(* IEC 61131-3 sources: PLC-IsaVODE/PLC-IsaVODE/samples/plc-programs (part 8) *)

(* ---- 638-IRTRANS_SERVER.ST ---- *)
TYPE

  oscat_NW_BUF_SHORT : ARRAY [0..1407] OF BYTE;
  oscat_NW_BUF_LONG  : ARRAY [0..4095] OF BYTE;

  oscat_NETWORK_BUFFER_SHORT :
  STRUCT
    SIZE   : UINT;
    BUFFER : oscat_NW_BUF_SHORT;
  END_STRUCT;

  oscat_NETWORK_BUFFER :
  STRUCT
    SIZE   : UINT;
    BUFFER : oscat_NW_BUF_LONG;
  END_STRUCT;

END_TYPE

TYPE
  oscat_IP_FIFO128_DATA  : ARRAY [1..128] OF BYTE;
  oscat_Mailbox  : ARRAY [1..16] OF BYTE;

  oscat_IP_FIFO_DATA :
  STRUCT
	X       : oscat_IP_FIFO128_DATA; (* IP_ID FIFO Speicher          *)
	Y       : oscat_IP_FIFO128_DATA; (* IP_ID Z�hler                 *)
	ID      : BYTE;                  (* h�chste vergabene id         *)
	MAX_ID  : BYTE;                  (* maximal Anmeldungen pro ID   *)
    INIT    : BOOL;                  (* Initialisierung durchgef�hrt *)
	EMPTY   : BOOL;                  (* FIFO leer                    *)
	FULL    : BOOL;                  (* FIFO voll                    *)
	TOP     : INT;                   (* maximale anzahl in FIFO      *)
	NW      : INT;                   (* Schreibzeiger                *)
	NR      : INT;                   (* Lesezeiger                   *)
  END_STRUCT;

  oscat_IP_C:
  STRUCT
  	C_MODE:			BYTE;          		(*W Mode: TCP/UCP AKTIV/PASSIV                               *)
	C_PORT:         WORD;          		(*W Portnummer                                               *)
	C_IP:           DWORD;         		(*W IP-Adresse gepackt wwxxyyzz = www.xxx.yyy.zzz            *)
    C_STATE:        BYTE;          		(*R Verbindungsstatus ON/OFF + Flanke ON/OFF                 *)
	C_ENABLE:       BOOL;          		(*W Freigabe f�r Connect                                     *)
    R_OBSERVE:      BOOL;          		(*W Empfang ueberwachen                                      *)
    TIME_RESET:     BOOL;          		(*W Alle Timer ruecksetzen                                   *)
	ERROR:          DWORD;         		(*R vvwwxxyy (vv = CON_ERROR, ww = SEN_ERROR, xx = REC_ERROR *)
    FIFO:           oscat_IP_FIFO_DATA; (*I IP FIFO Struktur                                         *)
	MAILBOX:		oscat_Mailbox;		(*I Mailbox: Datenbereich f�r Bausteindatenaustausch         *)
  END_STRUCT;
END_TYPE

FUNCTION_BLOCK IRTRANS_SERVER_Block

	VAR_INPUT
		UDP_TCP :	BOOL;
	END_VAR

	VAR_OUTPUT
		S_ENABLE :	BOOL;
		R_ENABLE :	BOOL;
		ERROR :	DWORD;
	END_VAR

	VAR_IN_OUT
		IP_C :	oscat_IP_C;
		S_BUF :	oscat_NETWORK_BUFFER;
		R_BUF :	oscat_NETWORK_BUFFER;
	END_VAR

	VAR
		t :	TON;
	END_VAR

	IF NOT IP_C.C_ENABLE THEN
		IP_C.C_PORT := WORD#0;
		IP_C.C_IP := DWORD#00;
		IP_C.C_MODE := SEL(UDP_TCP,BYTE#5,BYTE#4);
		IP_C.C_ENABLE := TRUE;
		IP_C.R_OBSERVE := FALSE;
		IP_C.TIME_RESET := TRUE;
		S_BUF.SIZE := UINT#0;
		R_BUF.SIZE := UINT#0;
	END_IF;

	R_ENABLE := IP_C.C_STATE > BYTE#127;
	S_ENABLE := R_ENABLE AND (IP_C.MAILBOX[1] > BYTE#0 OR IP_C.C_MODE <> BYTE#5);
	ERROR := IP_C.ERROR;

	t(IN:= IP_C.ERROR > DWORD#0, PT:=T#5s);
	IF t.Q THEN
		IP_C.TIME_RESET := TRUE;
	END_IF;

END_FUNCTION_BLOCK

PROGRAM program0
	VAR
		UDP_TCP :	BOOL;
		S_ENABLE :	BOOL;
		R_ENABLE :	BOOL;
		ERROR :	DWORD;
		IP_C :	oscat_IP_C;
		S_BUF :	oscat_NETWORK_BUFFER;
		R_BUF :	oscat_NETWORK_BUFFER;

		func_block : IRTRANS_SERVER_Block;
	END_VAR
	func_block.UDP_TCP := UDP_TCP;
	func_block.IP_C := IP_C;
	func_block.S_BUF := S_BUF;
	func_block.R_BUF := R_BUF;

	func_block();
	S_ENABLE  := func_block.S_ENABLE;
	R_ENABLE  := func_block.R_ENABLE;
	ERROR  := func_block.ERROR;
	IP_C  := func_block.IP_C;
	S_BUF  := func_block.S_BUF;
	R_BUF  := func_block.R_BUF;

END_PROGRAM

CONFIGURATION Config0

  	RESOURCE Res0 ON PLC
    	TASK task0(INTERVAL := T#20ms,PRIORITY := 0);
    	PROGRAM instance0 WITH task0 : program0;
  	END_RESOURCE

END_CONFIGURATION

(* ---- 639-FT_PDT1.ST ---- *)
FUNCTION _REAL_TO_UDINT:UDINT
  VAR_INPUT
    X :	REAL;
  END_VAR

  IF REAL_TO_UDINT(0.5) = UDINT#1 THEN
    _REAL_TO_UDINT := REAL_TO_UDINT(x);
  ELSIF X > 0.0 THEN
    _REAL_TO_UDINT := REAL_TO_UDINT(x+0.5);
  ELSIF X < 0.0 THEN
    _REAL_TO_UDINT := REAL_TO_UDINT(x-0.5);
  ELSE
    _REAL_TO_UDINT := UDINT#0;
  END_IF;
END_FUNCTION

FUNCTION REAL_TO_TIME2:TIME
	VAR_INPUT
		IN :	REAL;
	END_VAR

	REAL_TO_TIME2 := DINT_TO_TIME(UDINT_TO_DINT(_REAL_TO_UDINT(IN)));
END_FUNCTION

FUNCTION_BLOCK T_PLC_US_Block
	VAR_OUTPUT
		T_PLC_US :	UDINT;
	END_VAR

	VAR_EXTERNAL
		PLC_TICKS_PER_SEC :	INT;
		PLC_SYS_TICK_CNT :	DINT;
	END_VAR

	VAR
		debug :	BOOL;
		N :	INT;
		Offset :	UDINT;
		temp :	DWORD := DWORD#1;
		mode :	BOOL;
		faktor :	UDINT;
		init :	BOOL;
		v_plc_ticks_per_sec :	UDINT;
		base :	UDINT := UDINT#1000000;
	END_VAR

	IF init = FALSE THEN
		v_plc_ticks_per_sec := INT_TO_UDINT(PLC_TICKS_PER_SEC);
		IF v_plc_ticks_per_sec = UDINT#1024 THEN
			faktor := UDINT#1000;
			mode := FALSE;
		ELSIF v_plc_ticks_per_sec > UDINT#0 THEN
			IF v_plc_ticks_per_sec <= base THEN
				faktor := base / v_plc_ticks_per_sec;
				mode := FALSE;
			ELSE
				faktor := v_plc_ticks_per_sec / base;
				mode := TRUE;
			END_IF;
		ELSE
			faktor := UDINT#1;
		END_IF;
		init := TRUE;
	END_IF;

	IF mode THEN
		T_PLC_US := DINT_TO_UDINT(PLC_SYS_TICK_CNT) / faktor;
	ELSE
		T_PLC_US := DINT_TO_UDINT(PLC_SYS_TICK_CNT) * faktor;
	END_IF;

	IF debug THEN
		T_PLC_US := (DWORD_TO_UDINT(SHL(UDINT_TO_DWORD(T_PLC_US),N) OR SHL(temp,N)) - UDINT#1) + Offset;
	END_IF;
END_FUNCTION_BLOCK

FUNCTION_BLOCK FT_DERIV
	VAR_INPUT
		IN :	REAL;
		K :	REAL := 1.0;
		RUN :	BOOL := TRUE;
	END_VAR

	VAR_OUTPUT
		OUT :	REAL;
	END_VAR

	VAR
		old :	REAL;
		tx :	UDINT;
		last :	UDINT;
		init :	BOOL;
		tc :	REAL;
		T_PLC_US :	T_PLC_US_Block;
	END_VAR

	T_PLC_US();
	tx:= T_PLC_US.T_PLC_US;
	tc := UDINT_TO_REAL(tx - last);

	IF NOT init THEN
		init := TRUE;
		old := in;
	ELSIF run AND tc > 0.0 THEN
		out := (in - old) / tc * 1000000.0 * K;
		old := in;
	ELSE
		out := 0.0;
	END_IF;

	last := tx;

	T_PLC_US();
	tx:= T_PLC_US.T_PLC_US;

	IF NOT init THEN
		init := TRUE;
	ELSIF run AND tx - last > UDINT#0 THEN
		out := (in - old) / UDINT_TO_REAL(tx - last) * 1000000.0 * K;
	ELSE
		out := 0.0;
	END_IF;
	old := in;
	last := tx;
END_FUNCTION_BLOCK

FUNCTION_BLOCK FT_PT1

	VAR_INPUT
		IN :	REAL;
		T :	TIME;
		K :	REAL := 1.0;
	END_VAR

	VAR_OUTPUT
		OUT :	REAL;
	END_VAR

	VAR
		last :	UDINT;
		tx :	UDINT;
		init :	BOOL;
		T_PLC_US :	T_PLC_US_Block;
	END_VAR

	T_PLC_US();
	tx:= T_PLC_US.T_PLC_US;

	IF NOT init OR T = t#0s THEN
		init := TRUE;
		out := K * in;
	ELSE
		out := out + (in * K - out) * UDINT_TO_REAL(Tx - last) / TIME_TO_REAL(T) * 1.0E-3;
		IF ABS(out) < 1.0E-20 THEN out := 0.0; END_IF;
	END_IF;
	last := tx;
END_FUNCTION_BLOCK

FUNCTION_BLOCK FT_PDT1_Block

	VAR_INPUT
		IN :	REAL;
		KP :	REAL := 1.0;
		TV :	REAL := 1.0;
		T1 :	REAL := 1.0;
	END_VAR

	VAR_OUTPUT
		Y :	REAL;
	END_VAR

	VAR
		diff :	FT_DERIV;
		_TP :	FT_PT1;
	END_VAR

	diff(IN := IN, K := TV);

	_tp(in := diff.out, T := REAL_TO_TIME2(T1));

	Y := KP * (_tp.out + IN);

END_FUNCTION_BLOCK

PROGRAM program0
	VAR
		IN :	REAL;
		KP :	REAL := 1.0;
		TV :	REAL := 1.0;
		T1 :	REAL := 1.0;

		Y :	REAL;
		func_block : FT_PDT1_Block;
	END_VAR
	func_block.IN :=IN;
	func_block.KP :=KP;
	func_block.TV :=TV;
	func_block.T1 :=T1;
	func_block();
	Y := func_block.Y;
END_PROGRAM

CONFIGURATION Config0

	VAR_GLOBAL
		PLC_TICKS_PER_SEC :	INT;
		PLC_SYS_TICK_CNT :	DINT;
	END_VAR

	RESOURCE Res0 ON PLC
		TASK task0(INTERVAL := T#20ms,PRIORITY := 0);
		PROGRAM instance0 WITH task0 : program0;
	END_RESOURCE

END_CONFIGURATION

(* ---- 640-BOILER.ST ---- *)
FUNCTION_BLOCK BOILER_Block

	VAR_INPUT
		T_UPPER :	REAL;
		T_LOWER :	REAL;
		PRESSURE :	BOOL := TRUE;
		ENABLE :	BOOL := TRUE;
		REQ_1 :	BOOL;
		REQ_2 :	BOOL;
		BOOST :	BOOL;
		T_UPPER_MIN :	REAL := REAL#50.0;
		T_UPPER_MAX :	REAL := REAL#60.0;
		T_LOWER_ENABLE :	BOOL;
		T_LOWER_MAX :	REAL := REAL#60.0;
		T_REQUEST_1 :	REAL := REAL#70.0;
		T_REQUEST_2 :	REAL := REAL#50.0;
		T_REQUEST_HYS :	REAL := REAL#5.0;
		T_PROTECT_HIGH :	REAL := REAL#80.0;
		T_PROTECT_LOW :	REAL := REAL#10.0;
	END_VAR

	VAR_OUTPUT
		HEAT :	BOOL;
		ERROR :	BOOL;
		STATUS :	BYTE;
	END_VAR

	VAR
		edge :	BOOL;
		boost_mode :	BOOL;
		flag_0 :	BOOL;
		flag_1 :	BOOL;
		flag_2 :	BOOL;
	END_VAR

	IF t_upper > t_protect_high THEN
		status := BYTE#1;
		heat := FALSE;
		error := TRUE;
	ELSIF t_upper < t_protect_low THEN
		status := BYTE#2;
		heat := TRUE;
		error := TRUE;
	ELSIF t_lower > T_protect_high AND t_lower_enable THEN
		status := BYTE#3;
		heat := FALSE;
		error := TRUE;
	ELSIF t_lower < t_protect_low AND t_lower_enable THEN
		status := BYTE#4;
		heat := TRUE;
		error := TRUE;
	ELSIF NOT pressure THEN
		status := BYTE#5;
		heat := FALSE;
		error := TRUE;
	ELSIF req_1 OR req_2 OR enable OR boost THEN
		error := FALSE;

		IF boost AND NOT edge AND t_upper < t_upper_max THEN
			status := BYTE#101;
			heat := TRUE;
			boost_mode := TRUE;
		ELSIF enable AND t_upper < T_upper_min THEN
			status := BYTE#102;
			heat := TRUE;
		ELSIF req_1 AND t_upper < T_request_1 THEN
			status := BYTE#103;
			heat := TRUE;
		ELSIF req_2 AND t_upper < t_request_2 THEN
			status := BYTE#104;
			heat := TRUE;
		END_IF;

		IF heat THEN
			IF (enable OR boost_mode) THEN
				flag_0 := TRUE;
				IF T_lower_enable AND T_lower > T_lower_max THEN
					flag_0 := FALSE;
					boost_mode := FALSE;
				ELSIF NOT T_lower_enable AND T_upper > T_upper_max THEN
					flag_0 := FALSE;
					boost_mode := FALSE;
				END_IF;
			ELSE
				flag_0 := FALSE;
			END_IF;
			flag_1 := (req_1 AND T_upper > T_request_1 + T_request_hys) AND req_1;
			flag_2 := (req_2 AND T_upper > T_request_2 + T_request_hys) AND req_2;

			heat := flag_0 OR flag_1 OR flag_2;
			IF heat = FALSE THEN status := BYTE#100; END_IF;
		END_IF;
	ELSE
		status := BYTE#100;
		heat := FALSE;
		error := FALSE;
	END_IF;
	edge := boost;

END_FUNCTION_BLOCK

PROGRAM program0
	VAR
		T_UPPER :	REAL;
		T_LOWER :	REAL;
		PRESSURE :	BOOL := TRUE;
		ENABLE :	BOOL := TRUE;
		REQ_1 :	BOOL;
		REQ_2 :	BOOL;
		BOOST :	BOOL;
		T_UPPER_MIN :	REAL := REAL#50.0;
		T_UPPER_MAX :	REAL := REAL#60.0;
		T_LOWER_ENABLE :	BOOL;
		T_LOWER_MAX :	REAL := REAL#60.0;
		T_REQUEST_1 :	REAL := REAL#70.0;
		T_REQUEST_2 :	REAL := REAL#50.0;
		T_REQUEST_HYS :	REAL := REAL#5.0;
		T_PROTECT_HIGH :	REAL := REAL#80.0;
		T_PROTECT_LOW :	REAL := REAL#10.0;
		HEAT :	BOOL;
		ERROR :	BOOL;
		STATUS :	BYTE;

		func_block : BOILER_Block;
	END_VAR
	func_block.T_UPPER := T_UPPER;
	func_block.T_LOWER := T_LOWER;
	func_block.PRESSURE := PRESSURE ;
	func_block.ENABLE    := ENABLE    ;
	func_block.REQ_1 := REQ_1;
	func_block.REQ_2 := REQ_2;
	func_block.BOOST := BOOST ;
	func_block.T_UPPER_MIN := T_UPPER_MIN ;
	func_block.T_UPPER_MAX    := T_UPPER_MAX    ;
	func_block.T_LOWER_ENABLE := T_LOWER_ENABLE;
	func_block.T_LOWER_MAX := T_LOWER_MAX;
	func_block.T_REQUEST_1 := T_REQUEST_1 ;
	func_block.T_REQUEST_2 := T_REQUEST_2 ;
	func_block.T_REQUEST_HYS    := T_REQUEST_HYS    ;
	func_block.T_PROTECT_HIGH := T_PROTECT_HIGH;
	func_block.T_PROTECT_LOW := T_PROTECT_LOW;

	func_block();
	HEAT  := func_block.HEAT;
	ERROR  := func_block.ERROR;
	STATUS  := func_block.STATUS;
END_PROGRAM

CONFIGURATION Config0
	RESOURCE Res0 ON PLC
		TASK task0(INTERVAL := T#20ms,PRIORITY := 0);
		PROGRAM instance0 WITH task0 : program0;
	END_RESOURCE
END_CONFIGURATION

(* ---- 641-RMP_SOFT.ST ---- *)
FUNCTION TIME_TO_UDINT2:UDINT
	VAR_INPUT
		X :	TIME;
	END_VAR

	TIME_TO_UDINT2 := DINT_TO_UDINT(TIME_TO_DINT(X));
END_FUNCTION

FUNCTION_BLOCK T_PLC_MS_block
	VAR_OUTPUT
		T_PLC_MS :	UDINT;
	END_VAR

	VAR_EXTERNAL
		PLC_TICKS_PER_SEC :	INT;
		PLC_SYS_TICK_CNT :	DINT;
	END_VAR

	VAR
		debug :	BOOL;(*Debug-Mode ON / OFF*)
		N :	INT;(*Debug-Faktor*)
		Offset :	UDINT;(*Debug-Offset*)
		temp :	DWORD := DWORD#1;(*Debug-Offset*)
		mode :	BOOL;(*modus*)
		faktor :	UDINT;(*Systemtakt-Faktor*)
		init :	BOOL;
		v_plc_ticks_per_sec :	UDINT;
		base :	UDINT := UDINT#1000;
	END_VAR

	IF init = FALSE THEN
		v_plc_ticks_per_sec := INT_TO_UDINT(PLC_TICKS_PER_SEC);
		IF v_plc_ticks_per_sec = UDINT#1024 THEN
			faktor := UDINT#1;
			mode := FALSE;
		ELSIF v_plc_ticks_per_sec > UDINT#0 THEN
			IF v_plc_ticks_per_sec <= base THEN
				faktor := base / v_plc_ticks_per_sec;
				mode := FALSE;
			ELSE
				faktor := v_plc_ticks_per_sec / base;
				mode := TRUE;
			END_IF;
		ELSE
			faktor := UDINT#1;
		END_IF;
		init := TRUE;
	END_IF;

	IF mode THEN
		T_PLC_MS := DINT_TO_UDINT(PLC_SYS_TICK_CNT) / faktor;
	ELSE
		T_PLC_MS := DINT_TO_UDINT(PLC_SYS_TICK_CNT) * faktor;
	END_IF;

	IF debug THEN
		T_PLC_MS := (DWORD_TO_UDINT(SHL(UDINT_TO_DWORD(T_PLC_MS),N) OR SHL(temp,N)) - UDINT#1) + Offset;
	END_IF;
END_FUNCTION_BLOCK

FUNCTION FRMP_B:BYTE
	VAR_INPUT
		START :	BYTE;
		DIR :	BOOL;
		TD :	TIME;
		TR :	TIME;
	END_VAR

	IF TD < TR THEN
		FRMP_B := MIN(UDINT_TO_BYTE(DWORD_TO_UDINT(SHL(TIME_TO_DWORD(TD), 8)) / TIME_TO_UDINT2(TR)), SEL(DIR, START, USINT_TO_BYTE(USINT#255 - BYTE_TO_USINT(START))));
		IF DIR THEN
			FRMP_B := USINT_TO_BYTE(BYTE_TO_USINT(START) + BYTE_TO_USINT(FRMP_B));
		ELSE
			FRMP_B := USINT_TO_BYTE(BYTE_TO_USINT(START) - BYTE_TO_USINT(FRMP_B));
		END_IF;
	ELSE
		FRMP_B := SEL(DIR, BYTE#0, BYTE#255);
	END_IF;
END_FUNCTION

FUNCTION_BLOCK _RMP_B
	VAR_INPUT
		DIR :	BOOL;
		E :	BOOL := TRUE;
		TR :	TIME;
	END_VAR

	VAR_IN_OUT
		RMP :	BYTE;
	END_VAR

	VAR
		T_PLC_MS :	T_PLC_MS_block;
		tx :	TIME;
		tl :	TIME;
		tn :	TIME;
		init :	BOOL;
		last_dir :	BOOL;
		start :	BYTE;
	END_VAR

	T_PLC_MS();
	tx := UDINT_TO_TIME(T_PLC_MS.T_PLC_MS);

	IF E AND init AND (dir = last_dir) AND (RMP <> SEL(DIR, BYTE#0, BYTE#255)) AND TR = tn THEN
		RMP := FRMP_B(start, DIR, tx - tl, TR);
	ELSE
		init := TRUE;
		tl := tx;
		tn := tr;
		start := RMP;
	END_IF;
	last_dir := dir;
END_FUNCTION_BLOCK

FUNCTION_BLOCK RMP_SOFT_Block

	VAR_INPUT
		IN :	BOOL;
		VAL :	BYTE;
		PT_ON :	TIME := T#100ms;
		PT_OFF :	TIME := T#100ms;
	END_VAR

	VAR_OUTPUT
		OUT :	BYTE := BYTE#00;
	END_VAR

	VAR
		rmp :	_RMP_B;
		tmp :	BYTE;
	END_VAR

	tmp := SEL(in, BYTE#0, val);
	IF tmp > out THEN
		(* we need to ramp down *)
		rmp(dir := TRUE, E := TRUE, TR := PT_ON, RMP := out);
		out := rmp.RMP;
		(* make sure out does not surpass tmp *)
		out := MIN(out, tmp);
	ELSIF tmp < out THEN
		(* we need to ramp up *)
		rmp(dir := FALSE, E := TRUE, TR := PT_OFF, RMP := out);
		out := rmp.RMP;
		(* make sure out does not surpass tmp *)
		out := MAX(out, tmp);
	ELSE
		(* no ramp necessary *)
		rmp(E := FALSE, RMP := out);
		out := rmp.RMP;
	END_IF;

END_FUNCTION_BLOCK

PROGRAM program0
	VAR
		IN :	BOOL;
		VAL :	BYTE;
		PT_ON :	TIME;
		PT_OFF : TIME;

		OUT  :	BYTE;

		func_block : RMP_SOFT_Block;
	END_VAR
		func_block.IN := IN;
		func_block.VAL := VAL;
		func_block.PT_ON := PT_ON;
		func_block.PT_OFF := PT_OFF;
		func_block();
		OUT  := func_block.OUT ;

END_PROGRAM

CONFIGURATION Config0
	VAR_GLOBAL
		PLC_TICKS_PER_SEC :	INT;
		PLC_SYS_TICK_CNT :	DINT;
	END_VAR

  	RESOURCE Res0 ON PLC
    	TASK task0(INTERVAL := T#20ms,PRIORITY := 0);
    	PROGRAM instance0 WITH task0 : program0;
  	END_RESOURCE
END_CONFIGURATION

(* ---- 642-TUNE2.ST ---- *)
FUNCTION_BLOCK T_PLC_MS_block
	VAR_OUTPUT
		T_PLC_MS :	UDINT;
	END_VAR

	VAR_EXTERNAL
		PLC_TICKS_PER_SEC :	INT;
		PLC_SYS_TICK_CNT :	DINT;
	END_VAR

	VAR
		debug :	BOOL;(*Debug-Mode ON / OFF*)
		N :	INT;(*Debug-Faktor*)
		Offset :	UDINT;(*Debug-Offset*)
		temp :	DWORD := DWORD#1;(*Debug-Offset*)
		mode :	BOOL;(*modus*)
		faktor :	UDINT;(*Systemtakt-Faktor*)
		init :	BOOL;
		v_plc_ticks_per_sec :	UDINT;
		base :	UDINT := UDINT#1000;
	END_VAR

	IF init = FALSE THEN
		v_plc_ticks_per_sec := INT_TO_UDINT(PLC_TICKS_PER_SEC);
		IF v_plc_ticks_per_sec = UDINT#1024 THEN
			faktor := UDINT#1;
			mode := FALSE;
		ELSIF v_plc_ticks_per_sec > UDINT#0 THEN
			IF v_plc_ticks_per_sec <= base THEN
				faktor := base / v_plc_ticks_per_sec;
				mode := FALSE;
			ELSE
				faktor := v_plc_ticks_per_sec / base;
				mode := TRUE;
			END_IF;
		ELSE
			faktor := UDINT#1;
		END_IF;
		init := TRUE;
	END_IF;

	IF mode THEN
		T_PLC_MS := DINT_TO_UDINT(PLC_SYS_TICK_CNT) / faktor;
	ELSE
		T_PLC_MS := DINT_TO_UDINT(PLC_SYS_TICK_CNT) * faktor;
	END_IF;

	IF debug THEN
		T_PLC_MS := (DWORD_TO_UDINT(SHL(UDINT_TO_DWORD(T_PLC_MS),N) OR SHL(temp,N)) - UDINT#1) + Offset;
	END_IF;
END_FUNCTION_BLOCK

FUNCTION TIME_TO_UDINT2:UDINT
	VAR_INPUT
		X :	TIME;
	END_VAR

	TIME_TO_UDINT2 := DINT_TO_UDINT(TIME_TO_DINT(X));
END_FUNCTION

FUNCTION_BLOCK TUNE2_Block

	VAR_INPUT
		SET :	BOOL;
		SU :	BOOL;
		SD :	BOOL;
		FU :	BOOL;
		FD :	BOOL;
		RST :	BOOL;
		SS :	REAL := 0.1;
		FS :	REAL := 5.0;
		LIMIT_L :	REAL;
		LIMIT_H :	REAL := 100.0;
		RST_VAL :	REAL;
		SET_VAL :	REAL := 100.0;
		TR :	TIME := T#500ms;
		S1 :	REAL := 2.0;
		S2 :	REAL := 10.0;
	END_VAR

	VAR_OUTPUT
		Y :	REAL;
	END_VAR

	VAR
		tx :	UDINT;
		start :	UDINT;
		state :	INT;
		in :	BOOL;
		step2 :	REAL;
		speed :	REAL;
		Y_start :	REAL;
		T_PLC_MS :	T_PLC_MS_block;
	END_VAR

	T_PLC_MS();
	tx:= T_PLC_MS.T_PLC_MS;

	IF rst THEN
		Y := RST_val;
		state := 0;
	ELSIF set THEN
		Y := SET_val;
		state := 0;
	ELSIF state > 0 THEN
		CASE state OF
			1 :
				in := su;
			2 :
				in := sd;
			3 :
				in := fu;
			4 :
				in := fd;
		END_CASE;
		IF NOT in AND tx - start <= TIME_TO_UDINT2(TR) THEN
			Y := Y_start + step2;
			state := 0;
		ELSIF in AND tx - start >= TIME_TO_UDINT2(TR) THEN
			Y := Y_start + UDINT_TO_REAL(tx - start - TIME_TO_UDINT2(TR)) * speed;
		ELSIF NOT in THEN
			state := 0;
		END_IF;
	ELSIF su THEN
		state := 1;
		start := tx;
		step2 := ss;
		speed := s1 * 1.0E-3;
		Y_start := Y;
	ELSIF sd THEN
		state := 2;
		start := tx;
		step2 := -ss;
		speed := -s1 * 1.0E-3;
		Y_start := Y;
	ELSIF fu THEN
		state := 3;
		start := tx;
		step2 := fs;
		speed := s2 * 1.0E-3;
		y_start := Y;
	ELSIF fd THEN
		state := 4;
		start := tx;
		step2 := -fs;
		speed := -s2 * 1.0E-3;
		y_start := Y;
	END_IF;
END_FUNCTION_BLOCK

PROGRAM program0
  	VAR
		SET :	BOOL;
		SU :	BOOL;
		SD :	BOOL;
		FU :	BOOL;
		FD :	BOOL;
		RST :	BOOL;
		SS :	REAL;
		FS :	REAL;
		LIMIT_L :	REAL;
		LIMIT_H :	REAL;
		RST_VAL :	REAL;
		SET_VAL :	REAL;
		TR :	TIME ;
		S1 :	REAL;
		S2 :	REAL;
		Y :	REAL;
		func_block : TUNE2_Block;
  	END_VAR
	func_block.SET := SET;
	func_block.SU := SU;
	func_block.SD := SD;
	func_block.FU := FU;
	func_block.FD := FD;
	func_block.RST := RST;
	func_block.SS:= SS;
	func_block.FS := FS;
	func_block.LIMIT_L := LIMIT_L;
	func_block.LIMIT_H := LIMIT_H;
	func_block.RST_VAL := RST_VAL;
	func_block.SET_VAL := SET_VAL;
	func_block.TR := TR;
	func_block.S1 := S1;
	func_block.S2 := S2;
	func_block();
	Y := func_block.Y;
END_PROGRAM

CONFIGURATION Config0
	VAR_GLOBAL
		PLC_TICKS_PER_SEC :	INT;
		PLC_SYS_TICK_CNT :	DINT;
	END_VAR

	RESOURCE Res0 ON PLC
		TASK task0(INTERVAL := T#20ms,PRIORITY := 0);
		PROGRAM instance0 WITH task0 : program0;
	END_RESOURCE
END_CONFIGURATION

(* ---- 643-AIN1.ST ---- *)
FUNCTION_BLOCK AIN1

	VAR_INPUT
		IN :	DWORD;
		SIGN_BIT :	INT := 255;
		ERROR_BIT :	INT := 255;
		ERROR_CODE_EN :	BOOL := FALSE;
		ERROR_CODE :	DWORD;
		OVERFLOW_BIT :	INT := 255;
		OVERFLOW_CODE_EN :	BOOL;
		OVERFLOW_CODE :	DWORD;
		BIT_0 :	INT;
		BIT_N :	INT := 31;
		OUT_MIN :	REAL;
		OUT_MAX :	REAL := 10.0;
		CODE_MIN :	DWORD;
		CODE_MAX :	DWORD := DWORD#16#FFFFFFFF;
		ERROR_OUTPUT :	REAL;
		OVERFLOW_OUTPUT :	REAL := 10.0;
	END_VAR

	VAR_OUTPUT
		OUT :	REAL;
		SIGN :	BOOL;
		ERROR :	BOOL;
		OVERFLOW :	BOOL;
	END_VAR

	VAR
		tB :	DWORD;
	END_VAR

	error := ((SHR(in,error_bit) AND DWORD#16#0000_0001) = DWORD#1) OR (error_code_en AND error_code = in);
	IF error THEN
		out := error_output;
		RETURN;
	END_IF;

	tb := SHR(SHL(in, 31 - bit_N), 31 - bit_N + Bit_0);

	overflow := ((SHR(in,overflow_bit) AND DWORD#16#0000_0001) = DWORD#1) OR (overflow_code_en AND overflow_code = in) OR (tb < code_min OR tb > code_max);
	IF overflow THEN
		out := overflow_output;
		RETURN;
	END_IF;

	sign := (SHR(in,sign_bit) AND DWORD#16#0000_0001) = DWORD#1;

	out := (UDINT_TO_REAL(DWORD_TO_UDINT(tb) - DWORD_TO_UDINT(code_min)) * (out_max - out_min) / UDINT_TO_REAL(DWORD_TO_UDINT(code_max) - DWORD_TO_UDINT(code_min)) + out_min);
	IF sign THEN out := out * -1.0; END_IF;

	(* extract error bit *)
	error := ((SHR(in,error_bit) AND DWORD#16#0000_0001) = DWORD#1) OR (error_code_en AND error_code = in);
	IF error THEN
		out := error_output;
		RETURN;
	END_IF;

	(* strip off the data input *)
	tb := SHR(SHL(in, 31 - bit_N), 31 - bit_N + Bit_0);

	(* extract overflow bit *)
	overflow := ((SHR(in,overflow_bit) AND DWORD#16#0000_0001) = DWORD#1) OR (overflow_code_en AND overflow_code = in) OR (tb < code_min OR tb > code_max);
	IF overflow THEN
		out := overflow_output;
		RETURN;
	END_IF;

	(* extract sign bit *)
	sign := (SHR(in,sign_bit) AND DWORD#16#0000_0001) = DWORD#1;

	(* convert in to out *)
	out := (UDINT_TO_REAL(DWORD_TO_UDINT(tb) - DWORD_TO_UDINT(code_min)) * (out_max - out_min) / UDINT_TO_REAL(DWORD_TO_UDINT(code_max) - DWORD_TO_UDINT(code_min)) + out_min);
	IF sign THEN out := out * - 1.0; END_IF;

END_FUNCTION_BLOCK

PROGRAM program0
  VAR
	IN               :	DWORD;
	SIGN_BIT         :	INT ;
	ERROR_BIT        :	INT ;
	ERROR_CODE_EN    :	BOOL ;
	ERROR_CODE       :	DWORD;
	OVERFLOW_BIT     :	INT ;
	OVERFLOW_CODE_EN :	BOOL;
	OVERFLOW_CODE    :	DWORD;
	BIT_0            :	INT;
	BIT_N            :	INT;
	OUT_MIN          :	REAL;
	OUT_MAX          :	REAL ;
	CODE_MIN         :	DWORD;
	CODE_MAX         :	DWORD ;
	ERROR_OUTPUT     :	REAL;
	OVERFLOW_OUTPUT  :	REAL ;

	OUT      :	REAL;
	SIGN     :	BOOL;
	ERROR    :	BOOL;
	OVERFLOW :	BOOL;

	func_block : AIN1;
  END_VAR
	func_block.IN               :=IN              ;
	func_block.SIGN_BIT         :=SIGN_BIT        ;
	func_block.ERROR_BIT        :=ERROR_BIT       ;
	func_block.ERROR_CODE_EN    :=ERROR_CODE_EN   ;
	func_block.ERROR_CODE       :=ERROR_CODE      ;
	func_block.OVERFLOW_BIT     :=OVERFLOW_BIT    ;
	func_block.OVERFLOW_CODE_EN :=OVERFLOW_CODE_EN;
	func_block.OVERFLOW_CODE    :=OVERFLOW_CODE   ;
	func_block.BIT_0            :=BIT_0           ;
	func_block.BIT_N            :=BIT_N           ;
	func_block.OUT_MIN          :=OUT_MIN         ;
	func_block.OUT_MAX          :=OUT_MAX         ;
	func_block.CODE_MIN         :=CODE_MIN        ;
	func_block.CODE_MAX         :=CODE_MAX        ;
	func_block.ERROR_OUTPUT     :=ERROR_OUTPUT    ;
	func_block.OVERFLOW_OUTPUT  :=OVERFLOW_OUTPUT ;

	func_block();
	OUT     := func_block.OUT     ;
	SIGN    := func_block.SIGN    ;
	ERROR   := func_block.ERROR   ;
	OVERFLOW:= func_block.OVERFLOW;
END_PROGRAM

CONFIGURATION Config0
  RESOURCE Res0 ON PLC
    TASK task0(INTERVAL := T#20ms,PRIORITY := 0);
    PROGRAM instance0 WITH task0 : program0;
  END_RESOURCE
END_CONFIGURATION

(* ---- 644-TN_SC_VIEWPORT.ST ---- *)
TYPE
  bya_TN_CHAR:       	ARRAY [0..1919] OF BYTE;
  bya_TN_BACKUP:     	ARRAY [0..1919] OF BYTE;
  bya_TN_COLOR:      	ARRAY [0..1919] OF BYTE;
  bya_TN_Line_Update:	ARRAY [0..23]   OF BOOL;

  us_TN_SCREEN :
  STRUCT
		bya_CHAR:			bya_TN_CHAR;
		bya_COLOR:			bya_TN_COLOR;
		bya_BACKUP:			bya_TN_BACKUP;
		bya_Line_Update:	bya_TN_Line_Update;

		by_Input_Exten_Code:    BYTE;
		by_Input_ASCII_Code:    BYTE;
		bo_Input_ASCII_IsNum:   BOOL;
		in_Page_Number:        	INT;                (* aktive Seiten-Nr.              *)
		in_Cursor_X:           	INT;                (* Cursor X-Position              *)
		in_Cursor_Y:           	INT;                (* Cursor Y-Position              *)
		in_EOS_Offset:         	INT;                (* End of String Offset           *)
		by_Clear_Screen_Attr:  	BYTE;               (* Clear-Screen Attr              *)
		bo_Clear_Screen:       	BOOL;               (* Clear-Screen ausl�sen          *)
		bo_Modal_Dialog:       	BOOL;               (* Modaler Dialog ist aktiv       *)
		bo_Menue_Bar_Dialog:   	BOOL;               (* Menue Dialog ist aktiv         *)

  END_STRUCT;
END_TYPE

FUNCTION_BLOCK TN_SC_VIEWPORT_Block

  VAR
    FB_TN_SC_WRITE :	TN_SC_WRITE;
    FB_FIX :	FIX;
    FB_TON :	TON;
  END_VAR

  VAR
    in_index :	INT;
    in_Color :	INT;
    by_Attr :	BYTE;
    in_count :	INT;
  END_VAR

  VAR_IN_OUT
    Xus_LOG_VIEWPORT :	us_LOG_VIEWPORT;
    Xus_LOG_CONTROL :	us_LOG_CONTROL_80;
    Xus_TN_SCREEN :	us_TN_SCREEN;
  END_VAR

  VAR_INPUT
    Iin_X :	INT;
    Iin_Y :	INT;
    Iin_Width :	INT;
    Idw_ATTR_1 :	DWORD;
    Idw_ATTR_2 :	DWORD;
    Iti_TIME :	TIME;
  END_VAR

  IF Xus_LOG_VIEWPORT.UPDATE AND FB_TON.Q THEN

    Xus_LOG_VIEWPORT.UPDATE := FALSE;

    FOR in_count := 1 TO Xus_LOG_VIEWPORT.COUNT DO

      in_index := Xus_LOG_VIEWPORT.LINE_ARRAY[in_count];

    in_Color := DWORD_TO_INT(Xus_LOG_CONTROL.MSG_OPTION[in_index] AND DWORD#2#1111);

      CASE in_Color OF
        0..3: by_Attr := BYTE_OF_DWORD(Idw_ATTR_1,INT_TO_BYTE(in_Color));
        4..7: by_Attr := BYTE_OF_DWORD(Idw_ATTR_2,INT_TO_BYTE(in_Color));
      ELSE
      by_Attr := BYTE_OF_DWORD(Idw_ATTR_1,BYTE#0);
      END_CASE;

      FB_FIX.str := Xus_LOG_CONTROL.MSG[in_index];
      FB_FIX.L   := Iin_Width;
      FB_FIX.C   := BYTE#32;
      FB_FIX.M   := INT#00;
      FB_FIX();

      FB_TN_SC_WRITE.Iin_Y			:= Iin_Y + in_count - INT#01;
      FB_TN_SC_WRITE.Iin_X			:= Iin_X;
      FB_TN_SC_WRITE.Iby_ATTR			:= by_Attr;
      FB_TN_SC_WRITE.Ist_STRING		:= FB_FIX.FIX;
      FB_TN_SC_WRITE.Xus_TN_SCREEN	:= Xus_TN_SCREEN;
      FB_TN_SC_WRITE();
      Xus_TN_SCREEN := FB_TN_SC_WRITE.Xus_TN_SCREEN;

    END_FOR;

    FB_TON.IN := FALSE;
    FB_TON.PT := Iti_TIME;
    FB_TON();

  END_IF;

  FB_TON.IN := TRUE;
  FB_TON.PT := Iti_TIME;
  FB_TON();

END_FUNCTION_BLOCK

PROGRAM program0
	VAR
		Xus_LOG_VIEWPORT :	us_LOG_VIEWPORT;
    Xus_LOG_CONTROL :	us_LOG_CONTROL_80;
    Xus_TN_SCREEN :	us_TN_SCREEN;
    Iin_X :	INT;
    Iin_Y :	INT;
    Iin_Width :	INT;
    Idw_ATTR_1 :	DWORD;
    Idw_ATTR_2 :	DWORD;
    Iti_TIME :	TIME;

		func_block : TN_SC_VIEWPORT_Block;
	END_VAR
	func_block.Xus_LOG_VIEWPORT := Xus_LOG_VIEWPORT;
	func_block.Xus_LOG_CONTROL := Xus_LOG_CONTROL;
	func_block.Xus_TN_SCREEN := Xus_TN_SCREEN;
	func_block.Iin_X := Iin_X;
  func_block.Iin_Y := Iin_Y;
	func_block.Iin_Width := Iin_Width;
	func_block.Idw_ATTR_1 := Idw_ATTR_1;
	func_block.Idw_ATTR_2 := Idw_ATTR_2;
  func_block.Iti_TIME := Iti_TIME;

	func_block();
	Xus_LOG_VIEWPORT  := func_block.Xus_LOG_VIEWPORT;
  Xus_LOG_CONTROL  := func_block.Xus_LOG_CONTROL;
  Xus_TN_SCREEN  := func_block.Xus_TN_SCREEN;
END_PROGRAM

CONFIGURATION Config0
	RESOURCE Res0 ON PLC
		TASK task0(INTERVAL := T#20ms,PRIORITY := 0);
		PROGRAM instance0 WITH task0 : program0;
	END_RESOURCE
END_CONFIGURATION

(* ---- 645-DT_TO_SDT.ST ---- *)
TYPE oscat_SDT :
STRUCT
	YEAR : INT;
	MONTH : INT;
	DAY : INT;
	WEEKDAY : INT;
	HOUR : INT;
	MINUTE : INT;
	SECOND : INT;
	MS : INT;
END_STRUCT;
END_TYPE

FUNCTION DT_TO_DATE2:UDINT

	VAR_INPUT
		IN :	UDINT;
	END_VAR

	DT_TO_DATE2 := (IN / UDINT#86400) * UDINT#86400;
END_FUNCTION

FUNCTION YEAR_OF_DATE:INT
	VAR_INPUT
		IDATE :	UDINT;
	END_VAR

	YEAR_OF_DATE := UDINT_TO_INT((idate+UDINT#43200) / UDINT#31557600 + UDINT#1970);
END_FUNCTION

FUNCTION DAY_OF_WEEK:INT

	VAR_INPUT
		IDATE :	UDINT;
	END_VAR

	DAY_OF_WEEK := UDINT_TO_INT((idate / UDINT#86400 + UDINT#3) MOD UDINT#7) + INT#01;
END_FUNCTION

FUNCTION LEAP_OF_DATE:BOOL

	VAR_INPUT
		IDATE :	UDINT;
	END_VAR

	LEAP_OF_DATE := SHL(UDINT_TO_DWORD((idate + UDINT#43200) / UDINT#31557600), 30) = DWORD#16#80000000;
END_FUNCTION

FUNCTION DAY_OF_YEAR:INT
	VAR_INPUT
		IDATE :	UDINT;
	END_VAR

	DAY_OF_YEAR := UDINT_TO_INT(((idate) / UDINT#86400) MOD UDINT#1461);
	IF DAY_OF_YEAR > 729 THEN
		IF DAY_OF_YEAR > 1095 THEN DAY_OF_YEAR := DAY_OF_YEAR - 1095; ELSE DAY_OF_YEAR := DAY_OF_YEAR - 729; END_IF;
	ELSIF DAY_OF_YEAR > 364 THEN
		DAY_OF_YEAR := DAY_OF_YEAR - 364;
	ELSE
		DAY_OF_YEAR := DAY_OF_YEAR + 1;
	END_IF;
END_FUNCTION

FUNCTION MONTH_OF_DATE:INT

	VAR_INPUT
		IDATE :	UDINT;
	END_VAR

	MONTH_OF_DATE := DAY_OF_YEAR(idate);
	IF MONTH_OF_DATE < 32 THEN
		MONTH_OF_DATE := 1;
	ELSIF LEAP_OF_DATE((IDATE)) THEN
		MONTH_OF_DATE := (MONTH_OF_DATE * 53 + 1668) / 1623;
	ELSE
		MONTH_OF_DATE := (MONTH_OF_DATE * 53 + 1700) / 1620;
	END_IF;
END_FUNCTION

FUNCTION DAY_OF_MONTH:INT
	VAR_INPUT
		IDATE :	UDINT;
	END_VAR

	day_of_month := day_of_year(idate);

	IF leap_of_Date((idate)) THEN
		CASE day_of_month OF
			32..60	:	day_of_month := day_of_month - 31;
			61..91	:	day_of_month := day_of_month - 60;
			92..121 :	day_of_month := day_of_month - 91;
			122..152:	day_of_month := day_of_month - 121;
			153..182:	day_of_month := day_of_month - 152;
			183..213:	day_of_month := day_of_month - 182;
			214..244:	day_of_month := day_of_month - 213;
			245..274:	day_of_month := day_of_month - 244;
			275..305:	day_of_month := day_of_month - 274;
			306..335:	day_of_month := day_of_month - 305;
			336..366:	day_of_month := day_of_month - 335;
		END_CASE;
	ELSE
		CASE day_of_month OF
			32..59	:	day_of_month := day_of_month - 31;
			60..90	:	day_of_month := day_of_month - 59;
			91..120 :	day_of_month := day_of_month - 90;
			121..151:	day_of_month := day_of_month - 120;
			152..181:	day_of_month := day_of_month - 151;
			182..212:	day_of_month := day_of_month - 181;
			213..243:	day_of_month := day_of_month - 212;
			244..273:	day_of_month := day_of_month - 243;
			274..304:	day_of_month := day_of_month - 273;
			305..334:	day_of_month := day_of_month - 304;
			335..365:	day_of_month := day_of_month - 334;
		END_CASE;
	END_IF;
END_FUNCTION

FUNCTION _INT_TO_UDINT:UDINT
	VAR_INPUT
		IN :	INT;
	END_VAR

	_INT_TO_UDINT := DINT_TO_UDINT(INT_TO_DINT(IN));
END_FUNCTION

FUNCTION_BLOCK DT_TO_SDT

	VAR_INPUT
		DTI :	UDINT;
	END_VAR

	VAR_OUTPUT
		SDT :	oscat_SDT;
	END_VAR

	VAR
		tmp :	UDINT;
		tdt :	UDINT;
	END_VAR

	tmp := DT_TO_DATE2(dti);
	tdt := dti - tmp;
	SDT.YEAR := YEAR_OF_DATE(tmp);
	SDT.MONTH := MONTH_OF_DATE(tmp);
	SDT.DAY := DAY_OF_MONTH(tmp);
	SDT.WEEKDAY := DAY_OF_WEEK(tmp);
	SDT.SECOND := UDINT_TO_INT(tdt MOD UDINT#60);
	SDT.MINUTE := UDINT_TO_INT((tdt / UDINT#60) MOD UDINT#60);
	SDT.HOUR := UDINT_TO_INT(tdt / UDINT#3600);

END_FUNCTION_BLOCK

PROGRAM program0
  VAR
    LocalVar0 : UDINT;
	LocalOUT  : oscat_SDT;
	func_block : DT_TO_SDT;
  END_VAR
	func_block.DTI  := LocalVar0;
	func_block();
	LocalOUT := func_block.SDT;
END_PROGRAM

CONFIGURATION Config0
  RESOURCE Res0 ON PLC
    TASK task0(INTERVAL := T#20ms,PRIORITY := 0);
    PROGRAM instance0 WITH task0 : program0;
  END_RESOURCE
END_CONFIGURATION

(* ---- 646-AUTORUN.ST ---- *)
FUNCTION UDINT_TO_TIME2:TIME

	VAR_INPUT
		IN :	UDINT;
	END_VAR

	UDINT_TO_TIME2 := DINT_TO_TIME(UDINT_TO_DINT(IN));

END_FUNCTION

FUNCTION_BLOCK T_PLC_MS_block
	VAR_OUTPUT
		T_PLC_MS :	UDINT;
	END_VAR

	VAR_EXTERNAL
		PLC_TICKS_PER_SEC :	INT;
		PLC_SYS_TICK_CNT :	DINT;
	END_VAR

	VAR
		debug :	BOOL;(*Debug-Mode ON / OFF*)
		N :	INT;(*Debug-Faktor*)
		Offset :	UDINT;(*Debug-Offset*)
		temp :	DWORD := DWORD#1;(*Debug-Offset*)
		mode :	BOOL;(*modus*)
		faktor :	UDINT;(*Systemtakt-Faktor*)
		init :	BOOL;
		v_plc_ticks_per_sec :	UDINT;
		base :	UDINT := UDINT#1000;
	END_VAR

	IF init = FALSE THEN
		v_plc_ticks_per_sec := INT_TO_UDINT(PLC_TICKS_PER_SEC);
		IF v_plc_ticks_per_sec = UDINT#1024 THEN
			faktor := UDINT#1;
			mode := FALSE;
		ELSIF v_plc_ticks_per_sec > UDINT#0 THEN
			IF v_plc_ticks_per_sec <= base THEN
				faktor := base / v_plc_ticks_per_sec;
				mode := FALSE;
			ELSE
				faktor := v_plc_ticks_per_sec / base;
				mode := TRUE;
			END_IF;
		ELSE
			faktor := UDINT#1;
		END_IF;
		init := TRUE;
	END_IF;

	IF mode THEN
		T_PLC_MS := DINT_TO_UDINT(PLC_SYS_TICK_CNT) / faktor;
	ELSE
		T_PLC_MS := DINT_TO_UDINT(PLC_SYS_TICK_CNT) * faktor;
	END_IF;

	IF debug THEN
		T_PLC_MS := (DWORD_TO_UDINT(SHL(UDINT_TO_DWORD(T_PLC_MS),N) OR SHL(temp,N)) - UDINT#1) + Offset;
	END_IF;

END_FUNCTION_BLOCK

FUNCTION TIME_TO_UDINT2:UDINT
	VAR_INPUT
		X :	TIME;
	END_VAR

	TIME_TO_UDINT2 := DINT_TO_UDINT(TIME_TO_DINT(X));
END_FUNCTION

FUNCTION FRMP_B:BYTE
	VAR_INPUT
		START :	BYTE;
		DIR :	BOOL;
		TD :	TIME;
		TR :	TIME;
	END_VAR

	IF TD < TR THEN
		FRMP_B := MIN(UDINT_TO_BYTE(DWORD_TO_UDINT(SHL(TIME_TO_DWORD(TD), 8)) / TIME_TO_UDINT2(TR)), SEL(DIR, START, USINT_TO_BYTE(USINT#255 - BYTE_TO_USINT(START))));
		IF DIR THEN
			FRMP_B := USINT_TO_BYTE(BYTE_TO_USINT(START) + BYTE_TO_USINT(FRMP_B));
		ELSE
			FRMP_B := USINT_TO_BYTE(BYTE_TO_USINT(START) - BYTE_TO_USINT(FRMP_B));
		END_IF;
	ELSE
		FRMP_B := SEL(DIR, BYTE#0, BYTE#255);
	END_IF;
END_FUNCTION

FUNCTION_BLOCK _RMP_B
	VAR_INPUT
		DIR :	BOOL;
		E :	BOOL := TRUE;
		TR :	TIME;
	END_VAR

	VAR_IN_OUT
		RMP :	BYTE;
	END_VAR

	VAR
		T_PLC_MS :	T_PLC_MS_block;
		tx :	TIME;
		tl :	TIME;
		tn :	TIME;
		init :	BOOL;
		last_dir :	BOOL;
		start :	BYTE;
	END_VAR

	T_PLC_MS();
	tx := UDINT_TO_TIME(T_PLC_MS.T_PLC_MS);

	IF E AND init AND (dir = last_dir) AND (RMP <> SEL(DIR, BYTE#0, BYTE#255)) AND TR = tn THEN
		RMP := FRMP_B(start, DIR, tx - tl, TR);
	ELSE
		init := TRUE;
		tl := tx;
		tn := tr;
		start := RMP;
	END_IF;
	last_dir := dir;
END_FUNCTION_BLOCK

FUNCTION_BLOCK AUTORUN_Block

	VAR_INPUT
		IN :	BOOL;
		TEST :	BOOL;
		ARE :	BOOL := TRUE;
		TRUN :	TIME;
		TOFF :	TIME;
	END_VAR

	VAR_OUTPUT
		OUT :	BOOL;
		ARO :	BOOL;
	END_VAR

	VAR_IN_OUT
		ARX :	BOOL;
	END_VAR

	VAR
		timer :	_RMP_B;
		val :	BYTE;
	END_VAR

	IF TOFF > T#0s THEN
		timer(DIR:= OUT, TR := SEL(OUT, TOFF, TRUN), RMP := val);
		val := timer.RMP;
	ELSE
		val := BYTE#255;
	END_IF;

	IF (NOT ARX AND ARE AND val = BYTE#0) OR TEST THEN
		val := BYTE#0;
		ARO := TRUE;
		ARX := TRUE;
	ELSIF val = BYTE#255 AND ARO THEN
		ARO := FALSE;
		ARX := FALSE;
	END_IF;

	out := IN OR ARO;

END_FUNCTION_BLOCK

PROGRAM program0
	VAR
		IN :	BOOL;
		TEST :	BOOL;
		ARE :	BOOL := TRUE;
		TRUN :	TIME;
		TOFF :	TIME;
		OUT :	BOOL;
		ARO :	BOOL;
		func_block : AUTORUN_Block;
	END_VAR
	func_block.IN := IN;
	func_block.TEST := TEST;
	func_block.ARE := ARE ;
	func_block.TRUN := TRUN;
	func_block.TOFF := TOFF;
	func_block();
	OUT  := func_block.OUT;
	ARO  := func_block.ARO;
END_PROGRAM

CONFIGURATION Config0
	VAR_GLOBAL
		PLC_TICKS_PER_SEC :	INT;
		PLC_SYS_TICK_CNT :	DINT;
	END_VAR
  	RESOURCE Res0 ON PLC
    	TASK task0(INTERVAL := T#20ms,PRIORITY := 0);
    	PROGRAM instance0 WITH task0 : program0;
  	END_RESOURCE
END_CONFIGURATION

(* ---- 647-SHA1_STREAM.ST ---- *)
TYPE
  oscat_aB0_19	: ARRAY [0..19]	OF BYTE;
  oscat_aB0_63	: ARRAY [0..63]	OF BYTE;
  oscat_aDW0_4	: ARRAY [0..4] 	OF DWORD;
  oscat_sDW0_79	: ARRAY [0..79] OF DWORD;

END_TYPE

FUNCTION DWORD_OF_BYTE:DWORD
	VAR_INPUT
		B3 :	BYTE;
		B2 :	BYTE;
		B1 :	BYTE;
		B0 :	BYTE;
	END_VAR

	DWORD_OF_BYTE := SHL(SHL(SHL(BYTE_TO_DWORD(B3),8) OR BYTE_TO_DWORD(B2),8) OR BYTE_TO_DWORD(B1),8) OR BYTE_TO_DWORD(B0);

END_FUNCTION

FUNCTION_BLOCK SHA1_STREAM_Block

	VAR_IN_OUT
		MODE :	INT;
		BUF :	oscat_aB0_63;
		SHA1 :	oscat_aB0_19;
		SIZE :	UDINT;
	END_VAR

	VAR_OUTPUT
		POS :	UDINT;
	END_VAR

	VAR
		hash :	oscat_aDW0_4;
		end :	UDINT;
		block :	UDINT;
		pad_1 :	BOOL;
		w :	oscat_sDW0_79;
		n :	INT;
		n1 :	INT;
		n2 :	INT;
		n3 :	INT;
		n4 :	INT;
		a :	DWORD;
		b :	DWORD;
		c :	DWORD;
		d :	DWORD;
		e :	DWORD;
		f :	DWORD;
		k :	DWORD;
		x :	DWORD;
	END_VAR

	CASE MODE OF

	1:
		hash[0] := DWORD#16#67452301;
		hash[1] := DWORD#16#EFCDAB89;
		hash[2] := DWORD#16#98BADCFE;
		hash[3] := DWORD#16#10325476;
		hash[4] := DWORD#16#C3D2E1F0;

		FOR n := 16 TO 79 DO
			w[n] := DWORD#0;
		END_FOR;

		block := DWORD_TO_UDINT(SHR(UDINT_TO_DWORD(SIZE),6)) + BOOL_TO_UDINT((UDINT_TO_BYTE(SIZE) AND BYTE#16#3F) > BYTE#55);

		pad_1 := FALSE;
		POS := UDINT#0;
		End := SIZE;
		SIZE := MIN(UDINT#64,End);
		MODE := 2;

	2:	FOR n := UDINT_TO_INT(SIZE) TO 63 DO
			BUF[n] := BYTE#0;
		END_FOR;

		IF SIZE < UDINT#64 AND NOT pad_1 THEN
			BUF[SIZE] := BYTE#2#1000_0000;
			pad_1 := TRUE;
		END_IF;

		POS := POS + SIZE;
		SIZE := MIN(UDINT#64,End - POS);

		n := 0;
		FOR n4 := 0 TO 15 DO
			n1 := n + 1;
			n2 := n + 2;
			n3 := n + 3;
			w[n4] := DWORD_OF_BYTE(BUF[n],BUF[n1],BUF[n2],BUF[n3]);
			n := n + 4;
		END_FOR;

		IF block = UDINT#0 THEN
			w[15] := SHL(UDINT_TO_DWORD(End),3);
			MODE := 3;
		ELSE
			block := block - UDINT#1;
		END_IF;

		FOR n := 16 TO 79 DO
			n1 := n - 3;
			n2 := n - 8;
			n3 := n - 14;
			n4 := n - 16;
			w[n] := ROL(w[n1] XOR w[n2] XOR w[n3] XOR w[n4],1);
		END_FOR;

		a := hash[0];
		b := hash[1];
		c := hash[2];
		d := hash[3];
		e := hash[4];

		FOR n := 0 TO 79 DO
			IF n <= 19 THEN
				f := (b AND c) OR (NOT(b) AND d);
				k := DWORD#16#5A827999;
			ELSIF n <= 39 THEN
				f := b XOR c XOR d;
				k := DWORD#16#6ED9EBA1;
			ELSIF n <= 59 THEN
				f := (b AND c) OR (b AND d) OR (c AND d);
				k := DWORD#16#8F1BBCDC;
			ELSE
				f := b XOR c XOR d;
				k := DWORD#16#CA62C1D6;
			END_IF;

			x := UDINT_TO_DWORD(DWORD_TO_UDINT(ROL(a,5)) + DWORD_TO_UDINT(f) + DWORD_TO_UDINT(e) + DWORD_TO_UDINT(k) + DWORD_TO_UDINT(w[n]));
			e := d;
			d := c;
			c := ROL(b,30);
			b := a;
			a := x;
		END_FOR;

		hash[0] := UDINT_TO_DWORD(DWORD_TO_UDINT(hash[0]) + DWORD_TO_UDINT(a));
		hash[1] := UDINT_TO_DWORD(DWORD_TO_UDINT(hash[1]) + DWORD_TO_UDINT(b));
		hash[2] := UDINT_TO_DWORD(DWORD_TO_UDINT(hash[2]) + DWORD_TO_UDINT(c));
		hash[3] := UDINT_TO_DWORD(DWORD_TO_UDINT(hash[3]) + DWORD_TO_UDINT(d));
		hash[4] := UDINT_TO_DWORD(DWORD_TO_UDINT(hash[4]) + DWORD_TO_UDINT(e));

	END_CASE;

	IF MODE = 3 THEN
		n2 := 0;
		FOR n := 0 TO 4 DO
			FOR n1 := 0 TO 3 DO
				hash[n] := ROL(hash[n],8);
				SHA1[n2] := DWORD_TO_BYTE(hash[n]);
				n2 := n2 + 1;
			END_FOR;
		END_FOR;
	END_IF;

END_FUNCTION_BLOCK

PROGRAM program0
	VAR
		MODE :	INT;
		BUF :	oscat_aB0_63;
		SHA1 :	oscat_aB0_19;
		SIZE :	UDINT;
		POS :	UDINT;

		func_block : SHA1_STREAM_Block;
	END_VAR
	func_block.MODE := MODE;
	func_block.BUF := BUF;
	func_block.SHA1 := SHA1;
	func_block.SIZE := SIZE;

	func_block();
  	MODE  := func_block.MODE;
	BUF  := func_block.BUF;
	SHA1  := func_block.SHA1;
	SIZE  := func_block.SIZE;
	POS  := func_block.POS;
END_PROGRAM

CONFIGURATION Config0
	RESOURCE Res0 ON PLC
		TASK task0(INTERVAL := T#20ms,PRIORITY := 0);
		PROGRAM instance0 WITH task0 : program0;
	END_RESOURCE
END_CONFIGURATION

(* ---- 648-GEN_SIN.ST ---- *)
FUNCTION _REAL_TO_DWORD: DWORD

  VAR_INPUT
    X :	REAL;
  END_VAR

  IF REAL_TO_DWORD(0.5) = DWORD#1 THEN
    _REAL_TO_DWORD := REAL_TO_DWORD(x);
  ELSIF X > 0.0 THEN
    _REAL_TO_DWORD := REAL_TO_DWORD(x+0.5);
  ELSIF X < 0.0 THEN
    _REAL_TO_DWORD := REAL_TO_DWORD(x-0.5);
  ELSE
    _REAL_TO_DWORD := DWORD#0;
  END_IF;
END_FUNCTION

FUNCTION _DWORD_TO_REAL:REAL
	VAR_INPUT
		IN :	DWORD;
	END_VAR

	_DWORD_TO_REAL := UDINT_TO_REAL(DWORD_TO_UDINT(IN));

END_FUNCTION

FUNCTION MULTIME:TIME
	VAR_INPUT
		T :	TIME;
		M :	REAL;
	END_VAR

	multime := DWORD_TO_TIME(_REAL_TO_DWORD(_DWORD_TO_REAL(TIME_TO_DWORD(t))*M));
END_FUNCTION

FUNCTION UDINT_TO_TIME2:TIME

	VAR_INPUT
		IN :	UDINT;
	END_VAR

	UDINT_TO_TIME2 := DINT_TO_TIME(UDINT_TO_DINT(IN));

END_FUNCTION

FUNCTION_BLOCK T_PLC_MS_block
	VAR_OUTPUT
		T_PLC_MS :	UDINT;
	END_VAR

	VAR_EXTERNAL
		PLC_TICKS_PER_SEC :	INT;
		PLC_SYS_TICK_CNT :	DINT;
	END_VAR

	VAR
		debug :	BOOL;(*Debug-Mode ON / OFF*)
		N :	INT;(*Debug-Faktor*)
		Offset :	UDINT;(*Debug-Offset*)
		temp :	DWORD := DWORD#1;(*Debug-Offset*)
		mode :	BOOL;(*modus*)
		faktor :	UDINT;(*Systemtakt-Faktor*)
		init :	BOOL;
		v_plc_ticks_per_sec :	UDINT;
		base :	UDINT := UDINT#1000;
	END_VAR

	IF init = FALSE THEN
		v_plc_ticks_per_sec := INT_TO_UDINT(PLC_TICKS_PER_SEC);
		IF v_plc_ticks_per_sec = UDINT#1024 THEN
			faktor := UDINT#1;
			mode := FALSE;
		ELSIF v_plc_ticks_per_sec > UDINT#0 THEN
			IF v_plc_ticks_per_sec <= base THEN
				faktor := base / v_plc_ticks_per_sec;
				mode := FALSE;
			ELSE
				faktor := v_plc_ticks_per_sec / base;
				mode := TRUE;
			END_IF;
		ELSE
			faktor := UDINT#1;
		END_IF;
		init := TRUE;
	END_IF;

	IF mode THEN
		T_PLC_MS := DINT_TO_UDINT(PLC_SYS_TICK_CNT) / faktor;
	ELSE
		T_PLC_MS := DINT_TO_UDINT(PLC_SYS_TICK_CNT) * faktor;
	END_IF;

	IF debug THEN
		T_PLC_MS := (DWORD_TO_UDINT(SHL(UDINT_TO_DWORD(T_PLC_MS),N) OR SHL(temp,N)) - UDINT#1) + Offset;
	END_IF;

END_FUNCTION_BLOCK

FUNCTION TIME_TO_REAL1:REAL

	VAR_INPUT
		X :	TIME;
	END_VAR

	TIME_TO_REAL1 := UDINT_TO_REAL(DINT_TO_UDINT(TIME_TO_DINT(X)));
END_FUNCTION

FUNCTION MODR : REAL
  VAR_INPUT
    IN : REAL;
    DIVI : REAL;
  END_VAR

  IF divi = 0.0 THEN
  	MODR := 0.0;
  ELSE
  	MODR := in - DINT_TO_REAL(FLOOR2(in / divi)) * divi;
  END_IF;
END_FUNCTION

FUNCTION FLOOR2 : DINT
  VAR_INPUT
    x : REAL;
  END_VAR

  FLOOR2 := REAL_TO_DINT(X);
  IF DINT_TO_REAL(FLOOR2) > X THEN
  	FLOOR2 := FLOOR2 - DINT#1;
  END_IF;
END_FUNCTION

FUNCTION SIGN_R : BOOL
  VAR_INPUT
    IN : REAL;
  END_VAR

  SIGN_R := in < 0.0;
END_FUNCTION

FUNCTION_BLOCK GEN_SIN_Block

	VAR_INPUT
		PT :	TIME;
		AM :	REAL := REAL#1.0;
		OS :	REAL;
		DL :	REAL;
	END_VAR

	VAR_OUTPUT
		Q :	BOOL;
		Out :	REAL;
	END_VAR

	VAR
		tx :	TIME;
		last :	TIME;
		init :	BOOL;
		temp :	REAL;
		T_PLC_MS :	T_PLC_MS_Block;
	END_VAR

	T_PLC_MS();
	tx:= UDINT_TO_TIME(T_PLC_MS.T_PLC_MS) - last;

	DL := modR(dl,1.0);
	IF dl < 0.0 THEN dl := 1.0 - dl; END_IF;

	IF NOT init THEN
		init := TRUE;
		last := tx;
		tx := t#0s;
	END_IF;

	IF tx >= pt THEN
		last := last + pt;
		tx := tx - pt;
	END_IF;

	IF pt > t#0s THEN temp := SIN(6.283185307179586476 * TIME_TO_REAL1(tx + multime(pt, dl)) / TIME_TO_REAL(pt)); END_IF;
	out := am * 0.5 *  temp + os;

	q := NOT sign_R(temp);

END_FUNCTION_BLOCK

PROGRAM program0
  VAR
	PT :	TIME := T#1s;
	AM :	REAL := REAL#1.0;
	OS :	REAL;
	DL :	REAL;
	Q :	BOOL;
	OUT :	REAL;
	func_block : GEN_SIN_Block;
  END_VAR
	func_block.PT  :=PT;
	func_block.AM  :=AM;
	func_block.OS  :=OS;
	func_block.DL  :=DL;
	func_block();
	Q := func_block.Q;
	OUT := func_block.OUT;
END_PROGRAM

CONFIGURATION Config0
	VAR_GLOBAL
		PLC_TICKS_PER_SEC :	INT;
		PLC_SYS_TICK_CNT :	DINT;
	END_VAR
	RESOURCE Res0 ON PLC
		TASK task0(INTERVAL := T#20ms,PRIORITY := 0);
		PROGRAM instance0 WITH task0 : program0;
	END_RESOURCE
END_CONFIGURATION

(* ---- 649-ACTUATOR_UD.ST ---- *)
FUNCTION_BLOCK T_PLC_MS_block
	VAR_OUTPUT
		T_PLC_MS :	UDINT;
	END_VAR

	VAR_EXTERNAL
		PLC_TICKS_PER_SEC :	INT;
		PLC_SYS_TICK_CNT :	DINT;
	END_VAR

	VAR
		debug :	BOOL;(*Debug-Mode ON / OFF*)
		N :	INT;(*Debug-Faktor*)
		Offset :	UDINT;(*Debug-Offset*)
		temp :	DWORD := DWORD#1;(*Debug-Offset*)
		mode :	BOOL;(*modus*)
		faktor :	UDINT;(*Systemtakt-Faktor*)
		init :	BOOL;
		v_plc_ticks_per_sec :	UDINT;
		base :	UDINT := UDINT#1000;
	END_VAR

	IF init = FALSE THEN
		v_plc_ticks_per_sec := INT_TO_UDINT(PLC_TICKS_PER_SEC);
		IF v_plc_ticks_per_sec = UDINT#1024 THEN
			faktor := UDINT#1;
			mode := FALSE;
		ELSIF v_plc_ticks_per_sec > UDINT#0 THEN
			IF v_plc_ticks_per_sec <= base THEN
				faktor := base / v_plc_ticks_per_sec;
				mode := FALSE;
			ELSE
				faktor := v_plc_ticks_per_sec / base;
				mode := TRUE;
			END_IF;
		ELSE
			faktor := UDINT#1;
		END_IF;
		init := TRUE;
	END_IF;

	IF mode THEN
		T_PLC_MS := DINT_TO_UDINT(PLC_SYS_TICK_CNT) / faktor;
	ELSE
		T_PLC_MS := DINT_TO_UDINT(PLC_SYS_TICK_CNT) * faktor;
	END_IF;

	IF debug THEN
		T_PLC_MS := (DWORD_TO_UDINT(SHL(UDINT_TO_DWORD(T_PLC_MS),N) OR SHL(temp,N)) - UDINT#1) + Offset;
	END_IF;
END_FUNCTION_BLOCK

FUNCTION_BLOCK ACTUATOR_UD_Block

	VAR_INPUT
		UD :	BOOL;
		_ON :	BOOL;
		MANUAL :	BOOL;
		UP :	BOOL;
		DN :	BOOL;
		OFF :	BOOL;
		YUP_IN :	BOOL;
		YDN_IN :	BOOL;
		_TON :	TIME;
		TOFF :	TIME;
		OUT_RETURN :	BOOL;
	END_VAR

	VAR_OUTPUT
		YUP :	BOOL;
		YDN :	BOOL;
		STATUS :	BYTE;
	END_VAR

	VAR
		tx :	TIME;
		last :	TIME;
		init :	BOOL;
		T_PLC_MS :	T_PLC_MS_Block;
	END_VAR

	T_PLC_MS();
	tx:= UDINT_TO_TIME(T_PLC_MS.T_PLC_MS);

	IF NOT init THEN
		last := tx;
		init := TRUE;
	ELSIF off THEN
		Yup := FALSE;
		Ydn := FALSE;
		last := tx;
		status := BYTE#101;

	ELSIF ((Yup OR Ydn) AND tx - last < _TON) THEN RETURN;
	ELSIF NOT yup AND NOT ydn AND tx - last < toff THEN	RETURN;

	ELSIF manual THEN
		status := BYTE#102;
		IF yup AND NOT up OR ydn AND NOT dn THEN
			ydn := FALSE;
			yup := FALSE;
			last := tx;
		ELSIF UP AND NOT DN AND NOT OFF THEN
			Ydn := FALSE;
			Yup := TRUE;
			last := tx;
			status := BYTE#103;
		ELSIF DN AND NOT UP AND NOT OFF THEN
			Yup := FALSE;
			Ydn := TRUE;
			last := tx;
			status := BYTE#104;
		ELSE
			IF YUP OR YDN THEN LAST := tx; END_IF;
			Yup := FALSE;
			Ydn := FALSE;
		END_IF;

	ELSE
		IF yup AND NOT ud OR ydn AND UD THEN
			yup := FALSE;
			ydn := FALSE;
			last := tx;
		ELSIF Ud AND _ON AND NOT OFF THEN
			Ydn := FALSE;
			Yup := TRUE;
			last := tx;
			status := BYTE#111;

		ELSIF NOT UD AND _ON AND NOT OFF THEN
			Yup := FALSE;
			Ydn := TRUE;
			last := tx;
			status := BYTE#112;
		ELSE
			IF Yup OR Ydn THEN last := tx; END_IF;
			Yup := FALSE;
			Ydn := FALSE;
			status := BYTE#110;
		END_IF;
	END_IF;

	IF Ydn AND Yup_in AND out_return THEN
		Ydn := FALSE;
		status := BYTE#1;
	END_IF;
	IF Yup AND Ydn_in AND out_return THEN
		Yup := FALSE;
		status := BYTE#2;
	END_IF;

END_FUNCTION_BLOCK

PROGRAM program0
	VAR
		UD :	BOOL;
		_ON :	BOOL;
		MANUAL :	BOOL;
		UP :	BOOL;
		DN :	BOOL;
		OFF :	BOOL;
		YUP_IN :	BOOL;
		YDN_IN :	BOOL;
		_TON :	TIME;
		TOFF :	TIME;
		OUT_RETURN :	BOOL;
		YUP :	BOOL;
		YDN :	BOOL;
		STATUS :	BYTE;
		func_block : ACTUATOR_UD_Block;
	END_VAR
	func_block.UD := UD;
	func_block._ON := _ON;
	func_block.MANUAL := MANUAL ;
	func_block.UP := UP;
	func_block.DN := DN;
	func_block.OFF := OFF ;
	func_block.YUP_IN := YUP_IN;
	func_block.YDN_IN := YDN_IN;
	func_block._TON := _TON ;
	func_block.TOFF := TOFF;
	func_block.OUT_RETURN := OUT_RETURN;
	func_block();
	YUP  := func_block.YUP;
	YDN  := func_block.YDN;
	STATUS  := func_block.STATUS;
END_PROGRAM

CONFIGURATION Config0
	VAR_GLOBAL
		PLC_TICKS_PER_SEC :	INT;
		PLC_SYS_TICK_CNT :	DINT;
	END_VAR
  	RESOURCE Res0 ON PLC
    	TASK task0(INTERVAL := T#20ms,PRIORITY := 0);
    	PROGRAM instance0 WITH task0 : program0;
  	END_RESOURCE
END_CONFIGURATION

(* ---- 650-FADE.ST ---- *)
FUNCTION_BLOCK T_PLC_MS_block
	VAR_OUTPUT
		T_PLC_MS :	UDINT;
	END_VAR

	VAR_EXTERNAL
		PLC_TICKS_PER_SEC :	INT;
		PLC_SYS_TICK_CNT :	DINT;
	END_VAR

	VAR
		debug :	BOOL;(*Debug-Mode ON / OFF*)
		N :	INT;(*Debug-Faktor*)
		Offset :	UDINT;(*Debug-Offset*)
		temp :	DWORD := DWORD#1;(*Debug-Offset*)
		mode :	BOOL;(*modus*)
		faktor :	UDINT;(*Systemtakt-Faktor*)
		init :	BOOL;
		v_plc_ticks_per_sec :	UDINT;
		base :	UDINT := UDINT#1000;
	END_VAR

	IF init = FALSE THEN
		v_plc_ticks_per_sec := INT_TO_UDINT(PLC_TICKS_PER_SEC);
		IF v_plc_ticks_per_sec = UDINT#1024 THEN
			faktor := UDINT#1;
			mode := FALSE;
		ELSIF v_plc_ticks_per_sec > UDINT#0 THEN
			IF v_plc_ticks_per_sec <= base THEN
				faktor := base / v_plc_ticks_per_sec;
				mode := FALSE;
			ELSE
				faktor := v_plc_ticks_per_sec / base;
				mode := TRUE;
			END_IF;
		ELSE
			faktor := UDINT#1;
		END_IF;
		init := TRUE;
	END_IF;

	IF mode THEN
		T_PLC_MS := DINT_TO_UDINT(PLC_SYS_TICK_CNT) / faktor;
	ELSE
		T_PLC_MS := DINT_TO_UDINT(PLC_SYS_TICK_CNT) * faktor;
	END_IF;

	IF debug THEN
		T_PLC_MS := (DWORD_TO_UDINT(SHL(UDINT_TO_DWORD(T_PLC_MS),N) OR SHL(temp,N)) - UDINT#1) + Offset;
	END_IF;
END_FUNCTION_BLOCK

FUNCTION _WORD_TO_DINT:DINT
	VAR_INPUT
		IN :	WORD;
	END_VAR
	_WORD_TO_DINT := UINT_TO_DINT(WORD_TO_UINT(IN));
END_FUNCTION

FUNCTION TIME_TO_UDINT2:UDINT
	VAR_INPUT
		X :	TIME;
	END_VAR

	TIME_TO_UDINT2 := DINT_TO_UDINT(TIME_TO_DINT(X));
END_FUNCTION

FUNCTION_BLOCK _RMP_W

	VAR_INPUT
		DIR :	BOOL;
		E :	BOOL := TRUE;
		TR :	TIME;
	END_VAR

	VAR_IN_OUT
		RMP :	WORD;
	END_VAR

	VAR
		T_PLC_MS :	T_PLC_MS_block;
		tx :	UDINT;
		tl :	UDINT;
		ptesss :	DINT;
		init :	BOOL;
		last_dir :	BOOL;
	END_VAR

	T_PLC_MS();
	tx := T_PLC_MS.T_PLC_MS;
	IF E AND init THEN
		(* we need to set tl = tx when direction changes *)
		IF dir XOR last_dir THEN
			tl := tx;
			last_dir := dir;
		END_IF;
		(* check_elapsed time and calculate only if necessary *)
		IF tr > t#0s THEN
			ptesss := DWORD_TO_DINT(UDINT_TO_DWORD(DWORD_TO_UDINT(SHL(UDINT_TO_DWORD(tx-tl), 16)) / TIME_TO_UDINT2(TR)));
		ELSE
			ptesss := DINT#65535;
		END_IF;
		IF ptesss > DINT#0 THEN
			(* perform the ptesss on the ramp *)
			tl := tx;
			(* calculate the ptesss response *)
			IF NOT dir THEN ptesss := - ptesss; END_IF;
			rmp := DINT_TO_WORD(LIMIT(DINT#0, _WORD_TO_DINT(rmp) + ptesss, DINT#65535));
		END_IF;
	ELSE
		tl := tx;
		init := TRUE;
	END_IF;
END_FUNCTION_BLOCK

FUNCTION_BLOCK RMP_W

	VAR_INPUT
		SET :	BOOL;
		PT :	TIME;
		E :	BOOL := TRUE;
		UP :	BOOL := TRUE;
		RST :	BOOL;
	END_VAR

	VAR_OUTPUT
		OUT :	WORD;
		BUSY :	BOOL;
		HIGH :	BOOL;
		LOW :	BOOL;
	END_VAR

	VAR
		rmp :	_RMP_W;
	END_VAR

	rmp(dir := UP, E := E, TR := PT, rmp := out);
	out := rmp.RMP;

	IF RST THEN
		out := WORD#0;
	ELSIF SET THEN
		out := WORD#65535;
	END_IF;

	low := out = WORD#0;
	high := out = WORD#65535;
	busy := NOT (low OR high) AND E;

END_FUNCTION_BLOCK

FUNCTION _WORD_TO_REAL:REAL
	VAR_INPUT
		IN :	WORD;
	END_VAR
	_WORD_TO_REAL := UINT_TO_REAL(WORD_TO_UINT(IN));
END_FUNCTION

FUNCTION_BLOCK FADE
	VAR_INPUT
		IN1 :	REAL;
		IN2 :	REAL;
		F :	BOOL;
		TF :	TIME;
		RST :	BOOL;
	END_VAR

	VAR_OUTPUT
		Y :	REAL;
	END_VAR

	VAR
		rmx :	RMP_W;
	END_VAR
	rmx(rst := rst AND NOT F, set := rst AND F, pt := TF, up := F);
	Y := (in2 - In1) / 65535.0 * _WORD_TO_REAL(rmx.out) + in1;

END_FUNCTION_BLOCK

PROGRAM program0
  VAR

	IN1 :	REAL;
	IN2 :	REAL;
	F   :	BOOL;
	TF  :	TIME;
	RST :	BOOL;

	Y :	REAL;

	func_block : FADE;
  END_VAR
	func_block.IN1 :=IN1;
	func_block.IN2 :=IN2;
	func_block.F   :=F  ;
	func_block.TF  :=TF ;
	func_block.RST :=RST;
	func_block();
	Y := func_block.Y;

END_PROGRAM

CONFIGURATION Config0
	VAR_GLOBAL
		PLC_TICKS_PER_SEC :	INT;
		PLC_SYS_TICK_CNT :	DINT;
	END_VAR
  	RESOURCE Res0 ON PLC
    	TASK task0(INTERVAL := T#20ms,PRIORITY := 0);
    	PROGRAM instance0 WITH task0 : program0;
  	END_RESOURCE
END_CONFIGURATION

(* ---- 651-FLOW_METER.ST ---- *)
FUNCTION_BLOCK T_PLC_MS_block
	VAR_OUTPUT
		T_PLC_MS :	UDINT;
	END_VAR

	VAR_EXTERNAL
		PLC_TICKS_PER_SEC :	INT;
		PLC_SYS_TICK_CNT :	DINT;
	END_VAR

	VAR
		debug :	BOOL;(*Debug-Mode ON / OFF*)
		N :	INT;(*Debug-Faktor*)
		Offset :	UDINT;(*Debug-Offset*)
		temp :	DWORD := DWORD#1;(*Debug-Offset*)
		mode :	BOOL;(*modus*)
		faktor :	UDINT;(*Systemtakt-Faktor*)
		init :	BOOL;
		v_plc_ticks_per_sec :	UDINT;
		base :	UDINT := UDINT#1000;
	END_VAR

	IF init = FALSE THEN
		v_plc_ticks_per_sec := INT_TO_UDINT(PLC_TICKS_PER_SEC);
		IF v_plc_ticks_per_sec = UDINT#1024 THEN
			faktor := UDINT#1;
			mode := FALSE;
		ELSIF v_plc_ticks_per_sec > UDINT#0 THEN
			IF v_plc_ticks_per_sec <= base THEN
				faktor := base / v_plc_ticks_per_sec;
				mode := FALSE;
			ELSE
				faktor := v_plc_ticks_per_sec / base;
				mode := TRUE;
			END_IF;
		ELSE
			faktor := UDINT#1;
		END_IF;
		init := TRUE;
	END_IF;

	IF mode THEN
		T_PLC_MS := DINT_TO_UDINT(PLC_SYS_TICK_CNT) / faktor;
	ELSE
		T_PLC_MS := DINT_TO_UDINT(PLC_SYS_TICK_CNT) * faktor;
	END_IF;

	IF debug THEN
		T_PLC_MS := (DWORD_TO_UDINT(SHL(UDINT_TO_DWORD(T_PLC_MS),N) OR SHL(temp,N)) - UDINT#1) + Offset;
	END_IF;
END_FUNCTION_BLOCK

FUNCTION_BLOCK INTEGRATE

	VAR_INPUT
		E :	BOOL := TRUE;
		X :	REAL;
		K :	REAL := 1.0;
	END_VAR

	VAR_IN_OUT
		Y :	REAL;
	END_VAR

	VAR
		X_last :	REAL;
		init :	BOOL;
		T_PLC_MS :	T_PLC_MS_block;
		last :	UDINT;
		tx :	UDINT;
	END_VAR

	T_PLC_MS();
	tx:= T_PLC_MS.T_PLC_MS;

	IF NOT init THEN
		init := TRUE;
		X_last := X;
	ELSIF E THEN
		Y := (X + X_LAST) * 0.5E-3 * UDINT_TO_REAL(tx-last) * K + Y;
		X_last := X;
	END_IF;
	last := tx;

END_FUNCTION_BLOCK

FUNCTION _INT_TO_UDINT:UDINT
	VAR_INPUT
		IN :	INT;
	END_VAR

	_INT_TO_UDINT := DINT_TO_UDINT(INT_TO_DINT(IN));
END_FUNCTION

FUNCTION FLOOR : INT
	VAR_INPUT
		x : REAL;
	END_VAR

	FLOOR := REAL_TO_INT(X);
	IF INT_TO_REAL(FLOOR) > X THEN
		floor := floor - 1;
	END_IF;
END_FUNCTION

FUNCTION_BLOCK FLOW_METER
	VAR_INPUT
		VX :	REAL;
		E :	BOOL;
		RST :	BOOL;
		PULSE_MODE :	BOOL;
		UPDATE_TIME :	TIME := T#1s;
	END_VAR

	VAR_OUTPUT
		F :	REAL;
	END_VAR

	VAR_IN_OUT
		X :	REAL;
		Y :	UDINT;
	END_VAR

	VAR
		T_PLC_MS :	T_PLC_MS_block;
		tx :	TIME;
		tl :	TIME;
		int1 :	INTEGRATE;
		init :	BOOL;
		e_last :	BOOL;
		tmp :	INT;
		x_last :	REAL;
		y_last :	UDINT;
	END_VAR

	IF NOT init THEN	(* init on power up *)
		init := TRUE;
		tl := tx;
		x_last := X;
		y_last := Y;
		int1.K := 2.7777777777777777E-4;
	END_IF;

	int1(E := NOT (RST OR PULSE_MODE) AND E, X := VX, Y := X);	(* gated operation *)
	X := int1.Y;

	IF RST THEN		(* reset *)
		X := 0.0;
		Y := UDINT#0;
		tl := tx;
		x_last := 0.0;
		y_last := UDINT#0;
	ELSIF E AND PULSE_MODE THEN	(* check for pulse mode *)
		IF NOT e_last THEN X := X + VX; END_IF;
	END_IF;
	e_last := E;

	(* reduce X to be less than 1 and increase Y respectively *)
	IF X > 1.0 THEN
		tmp := FLOOR(X);
		Y := Y + _INT_TO_UDINT(tmp);
		X := X - INT_TO_REAL(tmp);
	END_IF;

	(* calculate the current flow *)
	T_PLC_MS();
	tx := UDINT_TO_TIME(T_PLC_MS.T_PLC_MS);
	IF tx - tl >= UPDATE_TIME AND UPDATE_TIME > t#0s THEN
		F := (UDINT_TO_REAL(Y - y_last) + X - x_last) / TIME_TO_REAL(tx - tl) * 3.6E6;
		y_last := Y;
		x_last := X;
		tl := tx;
	END_IF;

END_FUNCTION_BLOCK

PROGRAM program0
  VAR
	VX :	REAL;
	E :	BOOL;
	RST :	BOOL;
	PULSE_MODE :	BOOL;
	UPDATE_TIME :	TIME := T#1s;

	F :	REAL;

	X :	REAL;
	Y :	UDINT;

	func_block : FLOW_METER;
  END_VAR
	func_block.VX:=VX;
	func_block.E:=E;
	func_block.RST:=RST;
	func_block.PULSE_MODE:=PULSE_MODE;
	func_block.UPDATE_TIME :=UPDATE_TIME ;
	func_block.X:=X;
	func_block.Y:=Y;
	func_block();
	F:= func_block.F;
	X:= func_block.X;
	Y:= func_block.Y;
END_PROGRAM

CONFIGURATION Config0
	VAR_GLOBAL
		PLC_TICKS_PER_SEC :	INT;
		PLC_SYS_TICK_CNT :	DINT;
	END_VAR
	RESOURCE Res0 ON PLC
		TASK task0(INTERVAL := T#20ms,PRIORITY := 0);
		PROGRAM instance0 WITH task0 : program0;
	END_RESOURCE
END_CONFIGURATION

(* ---- 652-BLIND_SHADE_S.ST ---- *)
TYPE
  oscat_STRING5               : STRING;
  oscat_STRING30              : STRING;
END_TYPE

TYPE oscat_CALENDAR :
	STRUCT
		UTC : UDINT;				(* world time UTC *)
		LDT : UDINT;				(* local time *)
		LDATE : UDINT;				(* local date *)
		LTOD : UDINT;				(* local time of day *)
		YEAR : INT;					(* year of LDATE *)
		MONTH : INT;				(* month of LDATE *)
		DAY : INT;					(* day of LDATE *)
		WEEKDAY : INT;				(* weekday of LDATE *)
		OFFSET : INT;				(* Time Zone Offset for Local time in minutes *)
		DST_EN : BOOL;				(* daylight savings time enable *)
		DST_ON : BOOL;				(* true when daylight savings time os on *)
		NAME : oscat_string5;		(* name of time zone *)
		LANGUAGE : INT;			    (* language number pls see language setup *)
		LONGITUDE : REAL;			(* longitude of current location *)
		LATITUDE : REAL;			(* latitude of current location *)
		SUN_RISE : UDINT;			(* sun_rise for current location *)
		SUN_SET : UDINT;			(* sun_set for current location *)
		SUN_MIDDAY : UDINT;			(* worldtime when sun stands at south position *)
		SUN_HEIGTH : REAL;			(* suns heigth at midday, south position *)
		SUN_HOR : REAL;				(* sun angle horizontal 0 = north in degrees *)
		SUN_VER : REAL;				(* sun angle vertical above horizon in degrees *)
		NIGHT : BOOL;				(* true between sun_set and sun_rise *)
		HOLIDAY : BOOL;				(* true when holiday *)
		HOLY_NAME : oscat_string30;	(* name of holiday *)
		WORK_WEEK : INT;			(* current work week *)
	END_STRUCT;
END_TYPE

FUNCTION DT_TO_TOD2:UDINT
	VAR_INPUT
		IN :	UDINT;
	END_VAR

	DT_TO_TOD2 := (IN MOD UDINT#86400) * UDINT#1000;
END_FUNCTION

FUNCTION TIME_TO_UDINT2:UDINT
	VAR_INPUT
		X :	TIME;
	END_VAR

	TIME_TO_UDINT2 := DINT_TO_UDINT(TIME_TO_DINT(X));
END_FUNCTION

FUNCTION_BLOCK BLIND_SHADE_S_Block

	VAR_INPUT
		UP :	BOOL;
		DN :	BOOL;
		S_IN :	BYTE;
		PI :	BYTE;
		ENABLE :	BOOL;
		SUN :	BOOL;
		HORZ1 :	REAL := 100.0;
		HORZ2 :	REAL := 260.0;
		VERT :	REAL := 90.0;
		ALERT :	BOOL;
		SUNRISE_OFFSET :	TIME := T#1h;
		SUNSET_PRESET :	TIME := T#1h;
		SHADE_DELAY :	TIME := T#60s;
		SHADE_POS :	BYTE;
		QU :	BOOL;
		QD :	BOOL;
		STATUS :	BYTE;
		PO :	BYTE;
	END_VAR

	VAR_IN_OUT
		CX :	oscat_CALENDAR;
	END_VAR

	VAR
		angle :	REAL;
		sun_delay :	TOF;
	END_VAR

	sun_delay(IN := sun, PT := shade_delay);

	IF ALERT THEN
	QU := TRUE;
	QD := FALSE;
	STATUS := BYTE#152;
	ELSIF UP AND DN AND ENABLE AND sun_delay.Q
	AND (CX.SUN_HOR > HORZ1) AND (CX.SUN_HOR < HORZ2)
	AND (CX.SUN_VER < VERT)
	AND (DT_TO_TOD2(CX.UTC) > CX.SUN_RISE + TIME_TO_UDINT2(sunrise_offset)) AND (DT_TO_TOD2(CX.UTC) < CX.SUN_SET - TIME_TO_UDINT2(sunset_preset)) THEN
	QU := UP;
	QD := DN;
	STATUS := BYTE#151;
	PO := MIN(PI, shade_pos);
	ELSE
	QU := UP;
	QD := DN;
	PO := PI;
	STATUS := S_IN;
	END_IF;

END_FUNCTION_BLOCK

PROGRAM program0
	VAR
		UP :	BOOL;
		DN :	BOOL;
		S_IN :	BYTE;
		PI :	BYTE;
		ENABLE :	BOOL;
		SUN :	BOOL;
		HORZ1 :	REAL := 100.0;
		HORZ2 :	REAL := 260.0;
		VERT :	REAL := 90.0;
		ALERT :	BOOL;
		SUNRISE_OFFSET :	TIME := T#1h;
		SUNSET_PRESET :	TIME := T#1h;
		SHADE_DELAY :	TIME := T#60s;
		SHADE_POS :	BYTE;
		QU :	BOOL;
		QD :	BOOL;
		STATUS :	BYTE;
		PO :	BYTE;
		CX :	oscat_CALENDAR;

		func_block : BLIND_SHADE_S_Block;
	END_VAR
	func_block.UP := UP;
	func_block.DN := DN;
	func_block.S_IN := S_IN ;
	func_block.PI    := PI    ;
	func_block.ENABLE := ENABLE;
	func_block.SUN := SUN;
	func_block.HORZ1 := HORZ1 ;
	func_block.HORZ2 := HORZ2 ;
	func_block.VERT    := VERT    ;
	func_block.ALERT := ALERT;
	func_block.SUNRISE_OFFSET := SUNRISE_OFFSET;
	func_block.SUNSET_PRESET := SUNSET_PRESET ;
	func_block.SHADE_DELAY := SHADE_DELAY ;
	func_block.SHADE_POS    := SHADE_POS    ;
	func_block.QU := QU;
	func_block.QD := QD;
	func_block.STATUS := STATUS ;
	func_block.PO := PO ;
	func_block.CX := CX ;

	func_block();
	CX  := func_block.CX;
END_PROGRAM

CONFIGURATION Config0
	RESOURCE Res0 ON PLC
		TASK task0(INTERVAL := T#20ms,PRIORITY := 0);
		PROGRAM instance0 WITH task0 : program0;
	END_RESOURCE
END_CONFIGURATION

(* ---- 653-IP2GEO.ST ---- *)
FUNCTION_BLOCK IP2GEO

  VAR_IN_OUT
    IP_C :	oscat_IP_C;
    S_BUF :	oscat_NETWORK_BUFFER;
    R_BUF :	oscat_NETWORK_BUFFER;
    GEO :	oscat_IP2GEO_DATA;
  END_VAR

  VAR_INPUT
    IP :	DWORD;
    ACTIVATE :	BOOL;
  END_VAR

  VAR_OUTPUT
    BUSY :	BOOL;
    DONE :	BOOL;
    ERROR_C :	DWORD;
    ERROR_T :	BYTE;
  END_VAR

  VAR
    CTRL :	oscat_XML_CONTROL;
    XML_READER :	XML_READER;
    URL_DATA :	oscat_url;
    DNS_CLIENT :	DNS_CLIENT;
    STRING_TO_URL :	STRING_TO_URL;
    HTTP_GET :	HTTP_GET;
    FLOAT_TO_REAL :	FLOAT_TO_REAL;
    last_state :	BOOL;
    value_int :	INT;
    value_real :	REAL;
    v_real :	REAL;
    state :	INT;
    IP4_TO_STRING :	IP4_TO_STRING;
    IP4_DECODE :	IP4_DECODE;
    CHK_REAL :	CHK_REAL;
  END_VAR

  CASE state OF

  00:
    IF ACTIVATE AND NOT last_state THEN
      state := 20;
    DONE := FALSE;
    BUSY := TRUE;
    ERROR_C := DWORD#0;
    ERROR_T := BYTE#0;
    END_IF;

  20:
    STRING_TO_URL.STR:='http://ipinfodb.com/ip_query.php?timezone=true&IP=';
    STRING_TO_URL.DEFAULT_PROTOCOL:='';
    STRING_TO_URL.DEFAULT_PATH:='';
    STRING_TO_URL();
    URL_DATA:=STRING_TO_URL.STRING_TO_URL;

    IF IP > DWORD#0 THEN
      IP4_TO_STRING(IP4:=IP);
      URL_DATA.QUERY := CONCAT(URL_DATA.QUERY,IP4_TO_STRING.IP4_TO_STRING);
    END_IF;

    state := 40;

  40:
    IF DNS_CLIENT.DONE THEN
      state := 60;
    ELSIF (DNS_CLIENT.ERROR > DWORD#00) THEN
      ERROR_C := DNS_CLIENT.ERROR;
    ERROR_T := BYTE#01;
      state   := 100;
    END_IF;

  60:
    IF HTTP_GET.DONE THEN
      state := 80;
      CTRL.START_POS := HTTP_GET.BODY_START;
      CTRL.STOP_POS  := HTTP_GET.BODY_STOP;
      CTRL.COMMAND   := WORD#2#10000000_00011000;
    CTRL.WATCHDOG  := T#1ms;

    ELSIF (HTTP_GET.ERROR > DWORD#00) THEN
      ERROR_C := HTTP_GET.ERROR;
      ERROR_T := BYTE#02;
      state   := 100;
    END_IF;

  80:
    XML_READER.CTRL := CTRL;
    XML_READER.BUF  := R_BUF.BUFFER;
    XML_READER();
    CTRL         := XML_READER.CTRL;
    R_BUF.BUFFER := XML_READER.BUF;

    IF CTRL.TYP < 98 THEN
      value_int := 0;
      value_real := 0.0;
      IF LEN(CTRL.VALUE) <= 20 THEN
            FLOAT_TO_REAL(FLT:=CTRL.VALUE);
        v_real :=FLOAT_TO_REAL.FLOAT_TO_REAL;
        CHK_REAL(X:= v_real);
        IF CHK_REAL.CHK_REAL = BYTE#0 THEN
          value_real := v_real;
          value_int := REAL_TO_INT(value_real);
        END_IF;
      END_IF;

      CASE UINT_TO_INT(CTRL.COUNT) OF

        07: IP4_DECODE(STR:=CTRL.VALUE);
            GEO.IP4 := IP4_DECODE.IP4_DECODE;
      10: GEO.STATE := EQ_STRING('OK',CTRL.VALUE);
      13: GEO.COUNTRY_CODE := CTRL.VALUE;
      16: GEO.COUNTRY_NAME := CTRL.VALUE;
      19: GEO.REGION_CODE := CTRL.VALUE;
      22: GEO.REGION_NAME := CTRL.VALUE;
      25: GEO.CITY := CTRL.VALUE;
      31: GEO.GEO_LATITUDE := value_real;
      34: GEO.GEO_LONGITUDE := value_real;
      37: GEO.TIME_ZONE_NAME := CTRL.VALUE;
      40: GEO.GMT_OFFSET := value_int;
      43: GEO.IS_DST := value_int > 0;
      END_CASE;

    ELSIF CTRL.TYP = 99 THEN
      DONE  := TRUE;
      state := 100;
    END_IF;

  100:
    IF (NOT HTTP_GET.DONE) THEN
      state := 0;
      BUSY  := FALSE;
      DONE := ERROR_T = BYTE#0;
    END_IF;

  END_CASE;

  DNS_CLIENT.IP_C     := IP_C;
  DNS_CLIENT.S_BUF    := S_BUF;
  DNS_CLIENT.R_BUF    := R_BUF;
  DNS_CLIENT.DOMAIN   := URL_DATA.DOMAIN;
  DNS_CLIENT.IP4_DNS  := DWORD#00;
  DNS_CLIENT.ACTIVATE := state=40;
  DNS_CLIENT();
  IP_C  := DNS_CLIENT.IP_C;
  S_BUF := DNS_CLIENT.S_BUF;
  R_BUF := DNS_CLIENT.R_BUF;

  HTTP_GET.IP_C        := IP_C;
  HTTP_GET.S_BUF       := S_BUF;
  HTTP_GET.R_BUF       := R_BUF;
  HTTP_GET.IP4         := DNS_CLIENT.IP4;
  HTTP_GET.GET         := state=60;
  HTTP_GET.MODE        := BYTE#2;
  HTTP_GET.UNLOCK_BUF  := state=100;
  HTTP_GET.URL_DATA    := URL_DATA;
  HTTP_GET();
  IP_C     := HTTP_GET.IP_C;
  S_BUF    := HTTP_GET.S_BUF;
  R_BUF    := HTTP_GET.R_BUF;
  URL_DATA := HTTP_GET.URL_DATA;

  last_state := ACTIVATE;

END_FUNCTION_BLOCK

(* ---- 654-DNS_CLIENT.ST ---- *)
FUNCTION_BLOCK DNS_CLIENT

	VAR

	END_VAR

	VAR_EXTERNAL

	END_VAR

	VAR
		IP4_DECODE :	IP4_DECODE;
		IP_FIFO :	IP_FIFO;
		CODE :	CODE;
		ip_state :	BYTE;
		ip_id :	BYTE;
		i :	INT;
		i1 :	INT;
		i2 :	INT;
		i3 :	INT;
		state :	INT;
		domain_copy :	STRING;
		activate_last :	BOOL;
		url_length :	INT;
		char :	BYTE;
		char_count :	INT;
		tid :	BYTE;
		anc :	INT;
		x :	BYTE;
		rr_stop :	BOOL;
		ttl_last :	DWORD;
		ttl_tmp :	DWORD;
		z :	INT;
	END_VAR

	VAR_IN_OUT
		IP_C :	oscat_IP_C;
		S_BUF :	oscat_NETWORK_BUFFER;
		R_BUF :	oscat_NETWORK_BUFFER;
	END_VAR

	VAR_INPUT
		ACTIVATE :	BOOL;
		DOMAIN :	STRING;
		IP4_DNS :	DWORD;
	END_VAR

	VAR_OUTPUT
		IP4 :	DWORD;
		DONE :	BOOL;
		ERROR :	DWORD;
	END_VAR

	CASE state OF

	00:	IF ACTIVATE AND NOT activate_last THEN
			DONE := FALSE;
			ERROR := DWORD#0;
			state := 5;
		END_IF;

	05:
		IP4_DECODE(str:=DOMAIN);
		IP4 := IP4_DECODE.IP4_DECODE;
		IF IP4 > DWORD#00 THEN
			DONE := TRUE;
			state := 0;
		ELSE
			ip_state := BYTE#1;
			ttl_last := DWORD#0;
			domain_copy := DOMAIN;
			state := 10;
		END_IF;

	10:	IF ip_state = BYTE#3 THEN
			url_length := LEN(domain_copy);
			char_count := 17 + url_length;
			FOR i := 0 TO char_count DO
				S_BUF.BUFFER[i] := BYTE#00;
			END_FOR;
			tid := UINT_TO_BYTE(BYTE_TO_UINT(tid) + UINT#1);
			S_BUF.BUFFER[01] := tid;
			S_BUF.BUFFER[02] := BYTE#16#01;
			S_BUF.BUFFER[05] := BYTE#16#01;
			i := url_length + 12;
			char_count := 0;
			WHILE i > 12 DO
				CODE(STR:=domain_copy,POS:=i - 12);
				char := CODE.CODE;
				IF char = BYTE#46 THEN
					S_BUF.BUFFER[i] := INT_TO_BYTE(char_count);
					char_count := 0;
				ELSE
					S_BUF.BUFFER[i] := char;
					char_count := char_count + 1;
				END_IF;
				i := i - 1;
			END_WHILE;
			S_BUF.BUFFER[i] := INT_TO_BYTE(char_count);
			i := url_length + 15;
			S_BUF.BUFFER[i] := BYTE#01;
			i := i + 2;
			S_BUF.BUFFER[i] := BYTE#01;
			i := i + 1;
			IP_C.C_PORT := WORD#53;
			IP_C.C_IP := IP4_DNS;
			IP_C.C_MODE := BYTE#1;
			IP_C.C_ENABLE := TRUE;
			IP_C.TIME_RESET := TRUE;
			IP_C.R_OBSERVE  := TRUE;
			S_BUF.SIZE := INT_TO_UINT(i);
			R_BUF.SIZE := UINT#0;
			state := 30;
		END_IF;

	30:	IF IP_C.ERROR <> DWORD#00 THEN
			ERROR := IP_C.ERROR;
			state := 99;

		ELSIF (S_BUF.SIZE = UINT#0) AND (tid = R_BUF.BUFFER[1]) AND (R_BUF.SIZE >= INT_TO_UINT(34 + url_length)) THEN
			ERROR := BYTE_TO_DWORD(R_BUF.BUFFER[3] AND BYTE#2#0000_1111);
			IF ERROR = DWORD#00 THEN
				anc := _BYTE_TO_INT(R_BUF.BUFFER[7]);
				IP_C.R_OBSERVE := FALSE;
				state := 40;
			ELSE
				state := 99;
			END_IF;
		END_IF;

	40:	IF anc > 0 THEN
			anc := anc - 1;
			z := UINT_TO_INT(R_BUF.SIZE);
			WHILE i < z DO
				x := R_BUF.BUFFER[i];
				IF rr_stop = FALSE THEN
					IF x > BYTE#63 THEN
						i := i + 1;
						rr_stop := TRUE;
					ELSIF x= BYTE#0 THEN
						rr_stop := TRUE;
					ELSE
						i := i + _BYTE_TO_INT(x);
					END_IF;
					i := i + 1;
				ELSE
					rr_stop := FALSE;
					i1 := i + 1;
					i3 := i + 3;
					IF R_BUF.BUFFER[i1] = BYTE#1 AND R_BUF.BUFFER[i3] = BYTE#1 THEN
						i := i + 4;
						i1 := i + 1;
						i2 := i + 2;
						i3 := i + 3;
						ttl_tmp := DWORD_OF_BYTE(R_BUF.BUFFER[i],R_BUF.BUFFER[i1],R_BUF.BUFFER[i2],R_BUF.BUFFER[i3]);
						i := i + 6;
						IF ttl_tmp >= ttl_last THEN
							ttl_last := ttl_tmp;
							i1 := i + 1;
							i2 := i + 2;
							i3 := i + 3;
							IP4 := DWORD_OF_BYTE(R_BUF.BUFFER[i],R_BUF.BUFFER[i1],R_BUF.BUFFER[i2],R_BUF.BUFFER[i3]);
						END_IF;
						i := i + 4;
					ELSE
						i := i + 9;
						i := i + _BYTE_TO_INT(R_BUF.BUFFER[i]) + 1;
					END_IF;
					EXIT;
				END_IF;
			END_WHILE;
		ELSE
			IF IP4 > DWORD#0 THEN
				DONE := TRUE;
			ELSE
				ERROR := DWORD#255;
			END_IF;
			state := 99;
		END_IF;

	99:	R_BUF.SIZE := UINT#0;
		ip_state := BYTE#4;
		state := 00;

	END_CASE;

	activate_last := ACTIVATE;

	IP_FIFO(FIFO:=IP_C.FIFO,STATE:=ip_state,ID:=ip_id);
	IP_C.FIFO:=IP_FIFO.FIFO;
	ip_state := IP_FIFO.STATE;
	ip_id:=IP_FIFO.ID;

END_FUNCTION_BLOCK

(* ---- 655-NET_VAR_CONTROL.ST ---- *)
TYPE
	oscat_nv_dw : ARRAY[1..8] OF DWORD;
END_TYPE

TYPE

	oscat_NW_BUF_LONG  : ARRAY [0..4095] OF BYTE;

	oscat_NETWORK_BUFFER :
	STRUCT
		SIZE   : UINT;
		BUFFER : oscat_NW_BUF_LONG;
	END_STRUCT;

END_TYPE

TYPE oscat_NET_VAR_DATA :
	STRUCT
		CYCLE : UDINT;
		STATE : BYTE;
		INDEX : INT;
		ID_MAX : USINT;
		ERROR_ID : BYTE;
		BUF_SIZE : UINT;
		S_BUF : oscat_NETWORK_BUFFER;
		R_BUF : oscat_NETWORK_BUFFER;
	END_STRUCT;
END_TYPE

FUNCTION_BLOCK NET_VAR_CONTROL_Block

	VAR_INPUT
		ACTIVATE :	BOOL;
		MASTER :	BOOL;
		UDP :	BOOL;
		REMOTE_IP4 :	DWORD;
		REMOTE_PORT :	WORD := WORD#10000;
		SCAN_TIME :	TIME := T#1s;
		WATCHDOG :	TIME := T#2s;
	END_VAR

	VAR_OUTPUT
		RUN :	BOOL;
		ERROR :	DWORD;
	END_VAR

	VAR_IN_OUT
		X :	oscat_NET_VAR_DATA;
	END_VAR

	VAR
		IPC :	IP_CONTROL;
		IP_C :	oscat_IP_C;
		step :	INT;
		activate_last :	BOOL;
		tscan :	TON;
		reset :	BOOL;
	END_VAR

	IF X.ERROR_ID > BYTE#0 THEN
		X.STATE := BYTE#0;
		ERROR := BYTE_TO_DWORD(X.ERROR_ID);
		X.ERROR_ID := BYTE#0;
		step := 999;
	END_IF;

	CASE step OF

	00:	IF ACTIVATE AND NOT activate_last OR reset THEN
			IF MASTER THEN
				IP_C.C_MODE := BYTE#0;
				step := 100;
			ELSE
				IP_C.C_MODE := BYTE#2;
				step := 200;
			END_IF;
			IF UDP THEN IP_C.C_MODE := IP_C.C_MODE OR BYTE#1; END_IF;

			IP_C.C_PORT := REMOTE_PORT;
			IP_C.C_IP := REMOTE_IP4;
			IP_C.TIME_RESET := TRUE;
			IP_C.C_ENABLE := TRUE;
			IP_C.R_OBSERVE := TRUE;
			X.S_BUF.SIZE := UINT#0;
			X.R_BUF.SIZE := UINT#0;
			X.CYCLE := UDINT#0;
			X.ERROR_ID := BYTE#0;
			reset := FALSE;
		END_IF;

	100:IF IP_C.C_STATE > BYTE#127 THEN
			X.STATE := BYTE#1;
			X.BUF_SIZE := UINT#4096;
			X.S_BUF.BUFFER[0] := UDINT_TO_BYTE(X.CYCLE);
			X.INDEX := 1;
			step := 110;
		END_IF;

	110:X.STATE := BYTE#0;
		X.S_BUF.SIZE := INT_TO_UINT(X.INDEX);
		step := 120;

	120:IF X.S_BUF.SIZE = UINT#0 AND X.R_BUF.SIZE >= UINT#1 THEN
			X.STATE := BYTE#2;
			X.BUF_SIZE := X.R_BUF.SIZE;
			X.INDEX := 1;
			X.ERROR_ID := BYTE#0;
			X.CYCLE := X.CYCLE + UDINT#1;
			ERROR := DWORD#0;
			RUN := TRUE;
			step := 130;
		END_IF;

	130:X.STATE := BYTE#0;
		X.R_BUF.SIZE := UINT#0;
		IF NOT ACTIVATE THEN
			step := 999;
		ELSIF tscan.Q THEN
			step := 100;
		END_IF;

	200:IF X.R_BUF.SIZE >= UINT#1 THEN
			X.STATE := BYTE#2;
			X.BUF_SIZE := X.R_BUF.SIZE;
			X.INDEX := 1;
			step := 210;
		END_IF;

	210:X.STATE := BYTE#1;
		X.BUF_SIZE := UINT#4096;
		X.S_BUF.BUFFER[0] := X.R_BUF.BUFFER[0];
		X.INDEX := 1;
		X.R_BUF.SIZE := UINT#0;
		step := 220;

	220:X.STATE := BYTE#0;
		X.S_BUF.SIZE := INT_TO_UINT(X.INDEX);
		step := 230;

	230:IF X.S_BUF.SIZE = UINT#0 THEN
			ERROR := DWORD#0;
			RUN := TRUE;
			IF NOT ACTIVATE THEN
				step := 999;
			ELSE
				step := 200;
			END_IF;
		END_IF;

	999:IP_C.C_ENABLE := FALSE;
		RUN := FALSE;
		step := 0;

	END_CASE;

	IPC(IP:= DWORD#0, PORT:= WORD#0 , TIME_OUT:= WATCHDOG, IP_C:= IP_C, S_BUF:= X.S_BUF, R_BUF:= X.R_BUF);
	X.R_BUF := IPC.R_BUF;
	X.S_BUF := IPC.S_BUF;
	IP_C    := IPC.IP_C;

	IF IP_C.ERROR > DWORD#0 THEN
		ERROR := IP_C.ERROR;
		RUN := FALSE;
		reset := TRUE;
		step := 0;
	END_IF;

	ACTIVATE_LAST := ACTIVATE;
	tscan(IN:= step <> 110 ,PT:=SCAN_TIME);

END_FUNCTION_BLOCK

PROGRAM program0
	VAR
		ACTIVATE :	BOOL;
		MASTER :	BOOL;
		UDP :	BOOL;
		REMOTE_IP4 :	DWORD;
		REMOTE_PORT :	WORD := WORD#10000;
		SCAN_TIME :	TIME := T#1s;
		WATCHDOG :	TIME := T#2s;
		RUN :	BOOL;
		ERROR :	DWORD;
		X :	oscat_NET_VAR_DATA;

		func_block : NET_VAR_CONTROL_Block;
	END_VAR
	func_block.ACTIVATE := ACTIVATE;
	func_block.MASTER := MASTER;
	func_block.UDP := UDP;
	func_block.REMOTE_IP4 := REMOTE_IP4;
	func_block.REMOTE_PORT := REMOTE_PORT;
	func_block.SCAN_TIME := SCAN_TIME;
	func_block.WATCHDOG := WATCHDOG;
	func_block.X := X;

	func_block();
  	RUN  := func_block.RUN;
	ERROR  := func_block.ERROR;
	X  := func_block.X;

END_PROGRAM

CONFIGURATION Config0
	RESOURCE Res0 ON PLC
		TASK task0(INTERVAL := T#20ms,PRIORITY := 0);
		PROGRAM instance0 WITH task0 : program0;
	END_RESOURCE
END_CONFIGURATION

(* ---- 656-ACTUATOR_PUMP.ST ---- *)
FUNCTION_BLOCK T_PLC_MS_block
	VAR_OUTPUT
		T_PLC_MS :	UDINT;
	END_VAR

	VAR_EXTERNAL
		PLC_TICKS_PER_SEC :	INT;
		PLC_SYS_TICK_CNT :	DINT;
	END_VAR

	VAR
		debug :	BOOL;(*Debug-Mode ON / OFF*)
		N :	INT;(*Debug-Faktor*)
		Offset :	UDINT;(*Debug-Offset*)
		temp :	DWORD := DWORD#1;(*Debug-Offset*)
		mode :	BOOL;(*modus*)
		faktor :	UDINT;(*Systemtakt-Faktor*)
		init :	BOOL;
		v_plc_ticks_per_sec :	UDINT;
		base :	UDINT := UDINT#1000;
	END_VAR

	IF init = FALSE THEN
		v_plc_ticks_per_sec := INT_TO_UDINT(PLC_TICKS_PER_SEC);
		IF v_plc_ticks_per_sec = UDINT#1024 THEN
			faktor := UDINT#1;
			mode := FALSE;
		ELSIF v_plc_ticks_per_sec > UDINT#0 THEN
			IF v_plc_ticks_per_sec <= base THEN
				faktor := base / v_plc_ticks_per_sec;
				mode := FALSE;
			ELSE
				faktor := v_plc_ticks_per_sec / base;
				mode := TRUE;
			END_IF;
		ELSE
			faktor := UDINT#1;
		END_IF;
		init := TRUE;
	END_IF;

	IF mode THEN
		T_PLC_MS := DINT_TO_UDINT(PLC_SYS_TICK_CNT) / faktor;
	ELSE
		T_PLC_MS := DINT_TO_UDINT(PLC_SYS_TICK_CNT) * faktor;
	END_IF;

	IF debug THEN
		T_PLC_MS := (DWORD_TO_UDINT(SHL(UDINT_TO_DWORD(T_PLC_MS),N) OR SHL(temp,N)) - UDINT#1) + Offset;
	END_IF;

END_FUNCTION_BLOCK

FUNCTION_BLOCK ONTIME_Block

	VAR_INPUT
		IN :	BOOL;
		RST :	BOOL;
	END_VAR

	VAR_IN_OUT
		SECONDS :	UDINT;
		CYCLES :	UDINT;
	END_VAR

	VAR
		tx :	UDINT;
		last :	UDINT;
		edge :	BOOL;
		init :	BOOL;
		ms :	UDINT;
		T_PLC_MS :	T_PLC_MS_Block;
	END_VAR

	T_PLC_MS();
	tx:= T_PLC_MS.T_PLC_MS;

	IF NOT init THEN
		init := TRUE;
		last := tx;
		ms := UDINT#0;
	END_IF;
	IF RST THEN
		SECONDS := UDINT#0;
		CYCLES := UDINT#0;
		last := tx;
		ms := UDINT#0;
	ELSIF IN THEN
		(* add the current milliseconds *)
		ms := (tx - last) + ms;
		IF ms >= UDINT#1000 THEN
			seconds := seconds + UDINT#1;
			ms := ms - UDINT#1000;
		END_IF;
		cycles := cycles + BOOL_TO_UDINT(NOT edge);
	END_IF;
	last := tx;
	edge := in;

END_FUNCTION_BLOCK

FUNCTION_BLOCK ACTUATOR_PUMP_Block

	VAR_INPUT
		IN :	BOOL;
		MANUAL :	BOOL;
		RST :	BOOL := FALSE;
		MIN_ONTIME :	TIME := T#10s;
		MIN_OFFTIME :	TIME := T#10s;
		RUN_EVERY :	TIME := T#10000m;
	END_VAR

	VAR_OUTPUT
		PUMP :	BOOL;
		RUNTIME :	UDINT;
		CYCLES :	UDINT;
	END_VAR

	VAR
		tx :	TIME;
		last_change :	TIME;
		meter :	ONTIME_Block;
		old_man :	BOOL;
		init :	BOOL;
		T_PLC_MS :	T_PLC_MS_Block;
	END_VAR

	T_PLC_MS();
	tx:= UDINT_TO_TIME(T_PLC_MS.T_PLC_MS);

	IF NOT init THEN
		init := TRUE;
		last_change := tx;
	ELSIF rst THEN
		rst := FALSE;
		runtime := UDINT#0;
		cycles := UDINT#0;
	ELSIF manual AND NOT pump AND NOT old_man THEN
		last_change := tx;
		pump := TRUE;
	ELSIF NOT manual AND old_man AND pump AND NOT in THEN
		last_change := tx;
		pump := FALSE;
	ELSIF in AND NOT pump AND tx - last_change >= min_offtime THEN
		last_change := tx;
		pump := TRUE;
	ELSIF pump AND NOT in AND NOT manual AND tx - last_change >= min_ontime THEN
		last_change := tx;
		pump := FALSE;
	ELSIF NOT pump AND (tx - last_change >= run_every) AND (run_every > T#0s) THEN
		last_change := tx;
		pump := TRUE;
	END_IF;

	meter(in := pump, SECONDS := runtime, CYCLES := cycles);
	cycles := meter.CYCLES;
	runtime := meter.SECONDS;

	old_man := manual;

END_FUNCTION_BLOCK

PROGRAM program0
	VAR
		IN :	BOOL;
		MANUAL :	BOOL;
		RST :	BOOL := FALSE;
		MIN_ONTIME :	TIME := T#10s;
		MIN_OFFTIME :	TIME := T#10s;
		RUN_EVERY :	TIME := T#10000m;
		PUMP :	BOOL;
		RUNTIME :	UDINT;
		CYCLES :	UDINT;
		func_block : ACTUATOR_PUMP_Block;
	END_VAR
	func_block.IN := IN;
	func_block.MANUAL := MANUAL;
	func_block.RST := RST ;
	func_block.MIN_ONTIME := MIN_ONTIME;
	func_block.MIN_OFFTIME := MIN_OFFTIME;
	func_block.RUN_EVERY := RUN_EVERY ;
	func_block();
	PUMP  := func_block.PUMP;
	RUNTIME  := func_block.RUNTIME;
	CYCLES  := func_block.CYCLES;
END_PROGRAM

CONFIGURATION Config0
	VAR_GLOBAL
		PLC_TICKS_PER_SEC :	INT;
		PLC_SYS_TICK_CNT :	DINT;
	END_VAR
  	RESOURCE Res0 ON PLC
    	TASK task0(INTERVAL := T#20ms,PRIORITY := 0);
    	PROGRAM instance0 WITH task0 : program0;
  	END_RESOURCE
END_CONFIGURATION

(* ---- 657-RDM.ST ---- *)
FUNCTION D_TRUNC : DINT
  VAR_INPUT
    x : REAL;
  END_VAR

  D_TRUNC := REAL_TO_DINT(X);
  IF X > 0.0 THEN
  	IF DINT_TO_REAL(D_TRUNC) > X THEN D_TRUNC := D_TRUNC - DINT#1; END_IF;
  ELSE
  	IF DINT_TO_REAL(D_TRUNC) < X THEN D_TRUNC := D_TRUNC + DINT#1; END_IF;
  END_IF;
END_FUNCTION

FUNCTION BIT_COUNT:INT

	VAR_INPUT
		IN :	DWORD;
	END_VAR

	VAR
		in_temp :	DWORD;
	END_VAR

	in_temp := IN;
	WHILE in_temp > DWORD#0 DO
		IF (in_temp AND DWORD#16#00000001) > DWORD#0 THEN Bit_Count := Bit_Count +1; END_IF;
		in_temp := SHR(in_temp,1);
	END_WHILE;

END_FUNCTION

FUNCTION FRACT:REAL
	VAR_INPUT
		X :	REAL;
	END_VAR

	IF ABS(x) < 2.0E9 THEN
		FRACT := x - DINT_TO_REAL(D_TRUNC(x));
	ELSE
		FRACT := 0.0;
	END_IF;

END_FUNCTION

FUNCTION_BLOCK T_PLC_MS_block
	VAR_OUTPUT
		T_PLC_MS :	UDINT;
	END_VAR

	VAR_EXTERNAL
		PLC_TICKS_PER_SEC :	INT;
		PLC_SYS_TICK_CNT :	DINT;
	END_VAR

	VAR
		debug :	BOOL;(*Debug-Mode ON / OFF*)
		N :	INT;(*Debug-Faktor*)
		Offset :	UDINT;(*Debug-Offset*)
		temp :	DWORD := DWORD#1;(*Debug-Offset*)
		mode :	BOOL;(*modus*)
		faktor :	UDINT;(*Systemtakt-Faktor*)
		init :	BOOL;
		v_plc_ticks_per_sec :	UDINT;
		base :	UDINT := UDINT#1000;
	END_VAR

	IF init = FALSE THEN
		v_plc_ticks_per_sec := INT_TO_UDINT(PLC_TICKS_PER_SEC);
		IF v_plc_ticks_per_sec = UDINT#1024 THEN
			faktor := UDINT#1;
			mode := FALSE;
		ELSIF v_plc_ticks_per_sec > UDINT#0 THEN
			IF v_plc_ticks_per_sec <= base THEN
				faktor := base / v_plc_ticks_per_sec;
				mode := FALSE;
			ELSE
				faktor := v_plc_ticks_per_sec / base;
				mode := TRUE;
			END_IF;
		ELSE
			faktor := UDINT#1;
		END_IF;
		init := TRUE;
	END_IF;

	IF mode THEN
		T_PLC_MS := DINT_TO_UDINT(PLC_SYS_TICK_CNT) / faktor;
	ELSE
		T_PLC_MS := DINT_TO_UDINT(PLC_SYS_TICK_CNT) * faktor;
	END_IF;

	IF debug THEN
		T_PLC_MS := (DWORD_TO_UDINT(SHL(UDINT_TO_DWORD(T_PLC_MS),N) OR SHL(temp,N)) - UDINT#1) + Offset;
	END_IF;

END_FUNCTION_BLOCK

FUNCTION BIT_LOAD_DW:DWORD

	VAR_INPUT
		IN :	DWORD;
		VAL :	BOOL;
		POS :	INT;
	END_VAR

	IF val THEN
		BIT_LOAD_DW := in OR SHL(DWORD#1,pos);
	ELSE
		BIT_LOAD_DW := in AND (NOT SHL(DWORD#1,pos));
	END_IF;

END_FUNCTION

FUNCTION BIT_OF_DWORD : BOOL
  VAR_INPUT
    IN : DWORD;
    N : INT;
  END_VAR

  BIT_OF_DWORD := (SHR(in,N) AND 16#00000001) > 0;
  (* from OSCAT library; www.oscat.de  *)
END_FUNCTION

FUNCTION _INT_TO_UDINT:UDINT
	VAR_INPUT
		IN :	INT;
	END_VAR

	_INT_TO_UDINT := DINT_TO_UDINT(INT_TO_DINT(IN));
END_FUNCTION

FUNCTION _DWORD_TO_REAL:REAL
	VAR_INPUT
		IN :	DWORD;
	END_VAR

	_DWORD_TO_REAL := UDINT_TO_REAL(DWORD_TO_UDINT(IN));

END_FUNCTION

FUNCTION_BLOCK RDM_block
	VAR_INPUT
		LAST :	REAL;
	END_VAR
	VAR_OUTPUT
		RDM :	REAL;
	END_VAR
	VAR
		T_PLC_MS :	T_PLC_MS_block;
		tn :	DWORD;
		tc :	INT;
	END_VAR
	T_PLC_MS();
	tn := UDINT_TO_DWORD(T_PLC_MS.T_PLC_MS);
	tc := Bit_Count(tn);

	tn:=BIT_LOAD_DW(tn,BIT_OF_DWORD(tn,2),31); (* tn.31 := tn.2; *)
	tn:=BIT_LOAD_DW(tn,BIT_OF_DWORD(tn,5),30); (* tn.30 := tn.5; *)
	tn:=BIT_LOAD_DW(tn,BIT_OF_DWORD(tn,4),29); (* tn.29 := tn.4; *)
	tn:=BIT_LOAD_DW(tn,BIT_OF_DWORD(tn,1),28); (* tn.28 := tn.1; *)
	tn:=BIT_LOAD_DW(tn,BIT_OF_DWORD(tn,0),27); (* tn.27 := tn.0; *)
	tn:=BIT_LOAD_DW(tn,BIT_OF_DWORD(tn,7),26); (* tn.26 := tn.7; *)
	tn:=BIT_LOAD_DW(tn,BIT_OF_DWORD(tn,6),25); (* tn.25 := tn.6; *)
	tn:=BIT_LOAD_DW(tn,BIT_OF_DWORD(tn,3),24); (* tn.24 := tn.3; *)

	tn := ROL(tn,Bit_Count(tn)) OR DWORD#16#80000001;
	tn := UDINT_TO_DWORD(DWORD_TO_UDINT(tn) MOD UDINT#71474513 + _INT_TO_UDINT(tc) + UDINT#77);
	RDM := fract(_DWORD_TO_REAL(tn) / 10000000.0 * (2.71828182845904523536028747135266249 - LIMIT_REAL(0.0,last,1.0)));
END_FUNCTION_BLOCK

PROGRAM program0
	VAR
	    LocalVar : REAL;
		LocalOUT  : REAL;
		func_block : RDM_block;
  	END_VAR
	func_block.LAST := LocalVar;
	func_block();
	LocalOUT := func_block.RDM;
END_PROGRAM

CONFIGURATION Config0
	VAR_GLOBAL
		PLC_TICKS_PER_SEC :	INT;
		PLC_SYS_TICK_CNT :	DINT;
	END_VAR

  	RESOURCE Res0 ON PLC
    	TASK task0(INTERVAL := T#20ms,PRIORITY := 0);
    	PROGRAM instance0 WITH task0 : program0;
  	END_RESOURCE
END_CONFIGURATION

(* ---- 658-GEN_SQR.ST ---- *)
FUNCTION UDINT_TO_TIME2:TIME

	VAR_INPUT
		IN :	UDINT;
	END_VAR

	UDINT_TO_TIME2 := DINT_TO_TIME(UDINT_TO_DINT(IN));

END_FUNCTION

FUNCTION_BLOCK T_PLC_MS_block
	VAR_OUTPUT
		T_PLC_MS :	UDINT;
	END_VAR

	VAR_EXTERNAL
		PLC_TICKS_PER_SEC :	INT;
		PLC_SYS_TICK_CNT :	DINT;
	END_VAR

	VAR
		debug :	BOOL;(*Debug-Mode ON / OFF*)
		N :	INT;(*Debug-Faktor*)
		Offset :	UDINT;(*Debug-Offset*)
		temp :	DWORD := DWORD#1;(*Debug-Offset*)
		mode :	BOOL;(*modus*)
		faktor :	UDINT;(*Systemtakt-Faktor*)
		init :	BOOL;
		v_plc_ticks_per_sec :	UDINT;
		base :	UDINT := UDINT#1000;
	END_VAR

	IF init = FALSE THEN
		v_plc_ticks_per_sec := INT_TO_UDINT(PLC_TICKS_PER_SEC);
		IF v_plc_ticks_per_sec = UDINT#1024 THEN
			faktor := UDINT#1;
			mode := FALSE;
		ELSIF v_plc_ticks_per_sec > UDINT#0 THEN
			IF v_plc_ticks_per_sec <= base THEN
				faktor := base / v_plc_ticks_per_sec;
				mode := FALSE;
			ELSE
				faktor := v_plc_ticks_per_sec / base;
				mode := TRUE;
			END_IF;
		ELSE
			faktor := UDINT#1;
		END_IF;
		init := TRUE;
	END_IF;

	IF mode THEN
		T_PLC_MS := DINT_TO_UDINT(PLC_SYS_TICK_CNT) / faktor;
	ELSE
		T_PLC_MS := DINT_TO_UDINT(PLC_SYS_TICK_CNT) * faktor;
	END_IF;

	IF debug THEN
		T_PLC_MS := (DWORD_TO_UDINT(SHL(UDINT_TO_DWORD(T_PLC_MS),N) OR SHL(temp,N)) - UDINT#1) + Offset;
	END_IF;

END_FUNCTION_BLOCK

FUNCTION MODR : REAL
  VAR_INPUT
    IN : REAL;
    DIVI : REAL;
  END_VAR

  IF divi = 0.0 THEN
  	MODR := 0.0;
  ELSE
  	MODR := in - DINT_TO_REAL(FLOOR2(in / divi)) * divi;
  END_IF;
END_FUNCTION

FUNCTION FLOOR2 : DINT
  VAR_INPUT
    x : REAL;
  END_VAR

  FLOOR2 := REAL_TO_DINT(X);
  IF DINT_TO_REAL(FLOOR2) > X THEN
  	FLOOR2 := FLOOR2 - DINT#1;
  END_IF;
END_FUNCTION

FUNCTION _REAL_TO_DWORD: DWORD

  VAR_INPUT
    X :	REAL;
  END_VAR

  IF REAL_TO_DWORD(0.5) = DWORD#1 THEN
    _REAL_TO_DWORD := REAL_TO_DWORD(x);
  ELSIF X > 0.0 THEN
    _REAL_TO_DWORD := REAL_TO_DWORD(x+0.5);
  ELSIF X < 0.0 THEN
    _REAL_TO_DWORD := REAL_TO_DWORD(x-0.5);
  ELSE
    _REAL_TO_DWORD := DWORD#0;
  END_IF;
END_FUNCTION

FUNCTION _DWORD_TO_REAL:REAL
	VAR_INPUT
		IN :	DWORD;
	END_VAR

	_DWORD_TO_REAL := UDINT_TO_REAL(DWORD_TO_UDINT(IN));

END_FUNCTION

FUNCTION MULTIME:TIME
	VAR_INPUT
		T :	TIME;
		M :	REAL;
	END_VAR

	multime := DWORD_TO_TIME(_REAL_TO_DWORD(_DWORD_TO_REAL(TIME_TO_DWORD(t))*M));
END_FUNCTION

FUNCTION_BLOCK GEN_SQR_Block

	VAR_INPUT
		PT :	TIME;
		AM :	REAL := REAL#1.0;
		OS :	REAL;
		DC :	REAL := REAL#0.5;
		DL :	REAL;
	END_VAR

	VAR_OUTPUT
		Q :	BOOL;
		Out :	REAL;
	END_VAR

	VAR
		tx :	TIME;
		last :	TIME;
		init :	BOOL;
		T_PLC_MS :	T_PLC_MS_Block;
	END_VAR

	IF dc = 0.0 THEN
		out := -am * 0.5 + os;
		Q := FALSE;
		RETURN;
	ELSIF dc = 1.0 THEN
		out := am * 0.5 + os;
		Q := TRUE;
		RETURN;
	END_IF;

	T_PLC_MS();
	tx:= UDINT_TO_TIME(T_PLC_MS.T_PLC_MS) - last;
	DL := modR(dl,1.0);
	IF dl < 0.0 THEN dl := 1.0 - dl; END_IF;
	dc := modR(dc,1.0);
	IF dc < 0.0 THEN dc := 1.0 - dc; END_IF;

	IF NOT init THEN
		init := TRUE;
		last := tx;
		tx := t#0s;
	END_IF;

	IF tx >= pt THEN
		last := last + pt;
		tx := tx - pt;
	END_IF;

	IF multime(pt, dl + dc) >= pt THEN
		IF tx >= multime(pt, dl + dc - 1.0) THEN
			out := -am * 0.5 + os;
			Q := FALSE;
		END_IF;
		IF tx >= multime(pt, dl) THEN
			out := am * 0.5 + os;
			Q := TRUE;
		END_IF;
	ELSE
		IF tx >= multime(pt, dl) THEN
			out := am * 0.5 + os;
			Q := TRUE;
		END_IF;
		IF tx >= multime(pt, dl + dc) THEN
			out := -am * 0.5 +os;
			Q := FALSE;
		END_IF;
	END_IF;

END_FUNCTION_BLOCK

PROGRAM program0
  VAR
	PT :	TIME;
	AM :	REAL := REAL#1.0;
	OS :	REAL;
	DC :	REAL := REAL#0.5;
	DL :	REAL;
	Q :	BOOL;
	Out :	REAL;
	func_block : GEN_SQR_Block;
  END_VAR
	func_block.PT  :=PT;
	func_block.AM  :=AM;
	func_block.OS  :=OS;
	func_block.DC  :=DC;
	func_block.DL  :=DL;
	func_block();
	Q := func_block.Q;
	OUT := func_block.OUT;
END_PROGRAM

CONFIGURATION Config0
	VAR_GLOBAL
		PLC_TICKS_PER_SEC :	INT;
		PLC_SYS_TICK_CNT :	DINT;
	END_VAR
	RESOURCE Res0 ON PLC
		TASK task0(INTERVAL := T#20ms,PRIORITY := 0);
		PROGRAM instance0 WITH task0 : program0;
	END_RESOURCE
END_CONFIGURATION

(* ---- 659-IRTRANS_DECODE.ST ---- *)
FUNCTION_BLOCK CHR_TO_STRING_Block
	VAR_INPUT
		C :	BYTE;
	END_VAR

	VAR_OUTPUT
		CHR_TO_STRING :	STRING;
	END_VAR

	CHR_TO_STRING := BYTE_TO_STRING(C);

END_FUNCTION_BLOCK

TYPE

  oscat_NW_BUF_SHORT : ARRAY [0..1407] OF BYTE;
  oscat_NW_BUF_LONG  : ARRAY [0..4095] OF BYTE;

  oscat_NETWORK_BUFFER_SHORT :
  STRUCT
    SIZE   : UINT;
    BUFFER : oscat_NW_BUF_SHORT;
  END_STRUCT;

  oscat_NETWORK_BUFFER :
  STRUCT
    SIZE   : UINT;
    BUFFER : oscat_NW_BUF_LONG;
  END_STRUCT;

END_TYPE

TYPE
  oscat_IP_FIFO128_DATA  : ARRAY [1..128] OF BYTE;
  oscat_Mailbox  : ARRAY [1..16] OF BYTE;

  oscat_IP_FIFO_DATA :
  STRUCT
	X       : oscat_IP_FIFO128_DATA; (* IP_ID FIFO Speicher          *)
	Y       : oscat_IP_FIFO128_DATA; (* IP_ID Z�hler                 *)
	ID      : BYTE;                  (* h�chste vergabene id         *)
	MAX_ID  : BYTE;                  (* maximal Anmeldungen pro ID   *)
    INIT    : BOOL;                  (* Initialisierung durchgef�hrt *)
	EMPTY   : BOOL;                  (* FIFO leer                    *)
	FULL    : BOOL;                  (* FIFO voll                    *)
	TOP     : INT;                   (* maximale anzahl in FIFO      *)
	NW      : INT;                   (* Schreibzeiger                *)
	NR      : INT;                   (* Lesezeiger                   *)
  END_STRUCT;

  oscat_IP_C:
  STRUCT
  	C_MODE:			BYTE;          		(*W Mode: TCP/UCP AKTIV/PASSIV                               *)
	C_PORT:         WORD;          		(*W Portnummer                                               *)
	C_IP:           DWORD;         		(*W IP-Adresse gepackt wwxxyyzz = www.xxx.yyy.zzz            *)
    C_STATE:        BYTE;          		(*R Verbindungsstatus ON/OFF + Flanke ON/OFF                 *)
	C_ENABLE:       BOOL;          		(*W Freigabe f�r Connect                                     *)
    R_OBSERVE:      BOOL;          		(*W Empfang ueberwachen                                      *)
    TIME_RESET:     BOOL;          		(*W Alle Timer ruecksetzen                                   *)
	ERROR:          DWORD;         		(*R vvwwxxyy (vv = CON_ERROR, ww = SEN_ERROR, xx = REC_ERROR *)
    FIFO:           oscat_IP_FIFO_DATA; (*I IP FIFO Struktur                                         *)
	MAILBOX:		oscat_Mailbox;		(*I Mailbox: Datenbereich f�r Bausteindatenaustausch         *)
  END_STRUCT;
END_TYPE

FUNCTION_BLOCK IRTRANS_DECODE_Block

	VAR_OUTPUT
		CMD :	BOOL;
		DEV :	STRING;
		KEY :	STRING;
		ERROR :	BOOL;
	END_VAR

	VAR_IN_OUT
		IP_C :	oscat_IP_C;
		R_BUF :	oscat_NETWORK_BUFFER;
	END_VAR

	VAR
		i :	INT;
		stop :	INT;
		received_string :	STRING;
		char :	STRING;
		CHR_TO_STRING :	CHR_TO_STRING_Block;
		z :	BYTE;
	END_VAR

	i := UINT_TO_INT(R_BUF.SIZE);
	IF i >= 5 AND (i <= 82) AND IP_C.MAILBOX[1] <> z THEN
		error := TRUE;
		i := i - 1;

		IF R_BUF.BUFFER[i] <> BYTE#10 THEN RETURN; END_IF;
		i := i - 1;
		IF R_BUF.BUFFER[i] <> BYTE#13 THEN RETURN; END_IF;
		i := i - 1;

		stop := 0;
		received_string := '';

		WHILE stop <= i DO
			CHR_TO_STRING(C:=R_BUF.BUFFER[stop]);
			char := CHR_TO_STRING.CHR_TO_STRING;
			received_string := CONCAT(received_string,char);
			stop := stop + INT#1;
		END_WHILE;

		stop := FIND(received_string,',');
		IF stop > 0 AND stop - 1 < i THEN
			DEV := LEFT(received_string,stop - 1);
			key := RIGHT(received_string,i - stop + 1);
			IF LEN(DEV) = 0 OR LEN(key) = 0 THEN RETURN; END_IF;
			cmd := TRUE;
			error := FALSE;
		END_IF;
	ELSE
		cmd := FALSE;
		error := FALSE;
	END_IF;

	z := IP_C.MAILBOX[1];

END_FUNCTION_BLOCK

PROGRAM program0
	VAR
		IP_C :	oscat_IP_C;
		R_BUF :	oscat_NETWORK_BUFFER;
		CMD :	BOOL;
		DEV :	STRING;
		KEY :	STRING;
		ERROR :	BOOL;

		func_block : IRTRANS_DECODE_Block;
	END_VAR
	func_block.IP_C := IP_C;
	func_block.R_BUF := R_BUF;

	func_block();
	IP_C  := func_block.IP_C;
	R_BUF  := func_block.R_BUF;
	CMD  := func_block.CMD;
	DEV  := func_block.DEV;
	KEY  := func_block.KEY;
	ERROR  := func_block.ERROR;

END_PROGRAM

CONFIGURATION Config0

  	RESOURCE Res0 ON PLC
    	TASK task0(INTERVAL := T#20ms,PRIORITY := 0);
    	PROGRAM instance0 WITH task0 : program0;
  	END_RESOURCE

END_CONFIGURATION

(* ---- 660-NET_VAR_BOOL8.ST ---- *)
TYPE

	oscat_NW_BUF_LONG  : ARRAY [0..4095] OF BYTE;

	oscat_NETWORK_BUFFER :
	STRUCT
		SIZE   : UINT;
		BUFFER : oscat_NW_BUF_LONG;
	END_STRUCT;

END_TYPE

TYPE oscat_NET_VAR_DATA :
	STRUCT
		CYCLE : UDINT;
		STATE : BYTE;
		INDEX : INT;
		ID_MAX : USINT;
		ERROR_ID : BYTE;
		BUF_SIZE : UINT;
		S_BUF : oscat_NETWORK_BUFFER;
		R_BUF : oscat_NETWORK_BUFFER;
	END_STRUCT;
END_TYPE

FUNCTION BIT_OF_DWORD : BOOL
  VAR_INPUT
    IN : DWORD;
    N : INT;
  END_VAR

  BIT_OF_DWORD := (SHR(in,N) AND 16#00000001) > 0;
END_FUNCTION

FUNCTION_BLOCK BYTE_TO_BITS_Block
	VAR_INPUT
		IN :	BYTE;
	END_VAR

	VAR_OUTPUT
		B0 :	BOOL;
		B1 :	BOOL;
		B2 :	BOOL;
		B3 :	BOOL;
		B4 :	BOOL;
		B5 :	BOOL;
		B6 :	BOOL;
		B7 :	BOOL;
	END_VAR

	B0 := BIT_OF_DWORD(BYTE_TO_DWORD(IN),0); (* IN.X0 *)
	B1 := BIT_OF_DWORD(BYTE_TO_DWORD(IN),1); (* IN.X1 *)
	B2 := BIT_OF_DWORD(BYTE_TO_DWORD(IN),2); (* IN.X2 *)
	B3 := BIT_OF_DWORD(BYTE_TO_DWORD(IN),3); (* IN.X3 *)
	B4 := BIT_OF_DWORD(BYTE_TO_DWORD(IN),4); (* IN.X4 *)
	B5 := BIT_OF_DWORD(BYTE_TO_DWORD(IN),5); (* IN.X5 *)
	B6 := BIT_OF_DWORD(BYTE_TO_DWORD(IN),6); (* IN.X6 *)
	B7 := BIT_OF_DWORD(BYTE_TO_DWORD(IN),7); (* IN.X7 *)
END_FUNCTION_BLOCK

FUNCTION BYTE_OF_BIT:BYTE
	VAR_INPUT
		B0 :	BOOL;
		B1 :	BOOL;
		B2 :	BOOL;
		B3 :	BOOL;
		B4 :	BOOL;
		B5 :	BOOL;
		B6 :	BOOL;
		B7 :	BOOL;
	END_VAR
	Byte_of_bit := SHL(SHL(SHL(SHL(SHL(SHL(SHL(BOOL_TO_BYTE(B7),1) OR BOOL_TO_BYTE(B6),1)
	OR BOOL_TO_BYTE(B5),1) OR BOOL_TO_BYTE(B4),1) OR BOOL_TO_BYTE(B3),1) OR BOOL_TO_BYTE(B2),1)
	OR BOOL_TO_BYTE(B1),1) OR BOOL_TO_BYTE(B0);
END_FUNCTION

FUNCTION_BLOCK NET_VAR_BOOL8_Block

	VAR_INPUT
		IN1 :	BOOL;
		IN2 :	BOOL;
		IN3 :	BOOL;
		IN4 :	BOOL;
		IN5 :	BOOL;
		IN6 :	BOOL;
		IN7 :	BOOL;
		IN8 :	BOOL;
	END_VAR

	VAR_OUTPUT
		OUT1 :	BOOL;
		OUT2 :	BOOL;
		OUT3 :	BOOL;
		OUT4 :	BOOL;
		OUT5 :	BOOL;
		OUT6 :	BOOL;
		OUT7 :	BOOL;
		OUT8 :	BOOL;
		ID :	BYTE;
	END_VAR

	VAR_IN_OUT
		X :	oscat_NET_VAR_DATA;
	END_VAR

	VAR
		init :	BOOL;
		index :	INT;
		index2 :	INT;
		_BYTE_TO_BITS :	BYTE_TO_BITS_Block;
	END_VAR

	IF NOT init THEN
		init := TRUE;
		X.ID_MAX := X.ID_MAX + USINT#1;
		ID := USINT_TO_BYTE(X.ID_MAX);
	END_IF;

	IF X.STATE > BYTE#0 AND X.ERROR_ID = BYTE#0 THEN
		index := X.index;
		IF INT_TO_UINT(index + 3) > X.BUF_SIZE THEN
			X.ERROR_ID := ID;
		ELSE
			IF X.STATE = BYTE#1 THEN
				X.S_BUF.BUFFER[index] := ID;
				index := index + 1;
				X.S_BUF.BUFFER[index] := BYTE#4;
				index := index + 1;
				X.S_BUF.BUFFER[index] := BYTE_OF_BIT(IN1,IN2,IN3,IN4,IN5,IN6,IN7,IN8);
				index := index + 1;

			ELSIF X.STATE = BYTE#2 THEN
				index2 := index + 1;
				IF X.R_BUF.BUFFER[index] <> ID OR X.R_BUF.BUFFER[index2] <> BYTE#4 THEN
					X.ERROR_ID := ID;
				ELSE
					index := index + 2;
					_BYTE_TO_BITS(IN:=X.R_BUF.BUFFER[index]);
					OUT1 := _BYTE_TO_BITS.B0;
					OUT2 := _BYTE_TO_BITS.B1;
					OUT3 := _BYTE_TO_BITS.B2;
					OUT4 := _BYTE_TO_BITS.B3;
					OUT5 := _BYTE_TO_BITS.B4;
					OUT6 := _BYTE_TO_BITS.B5;
					OUT7 := _BYTE_TO_BITS.B6;
					OUT8 := _BYTE_TO_BITS.B7;
					index := index + 1;
				END_IF;
			END_IF;
			X.index := index;
		END_IF;
	END_IF;

END_FUNCTION_BLOCK

PROGRAM program0
	VAR
		IN1 :	BOOL;
		IN2 :	BOOL;
		IN3 :	BOOL;
		IN4 :	BOOL;
		IN5 :	BOOL;
		IN6 :	BOOL;
		IN7 :	BOOL;
		IN8 :	BOOL;
		OUT1 :	BOOL;
		OUT2 :	BOOL;
		OUT3 :	BOOL;
		OUT4 :	BOOL;
		OUT5 :	BOOL;
		OUT6 :	BOOL;
		OUT7 :	BOOL;
		OUT8 :	BOOL;
		ID :	BYTE;
		X :	oscat_NET_VAR_DATA;

		func_block : NET_VAR_BOOL8_Block;
	END_VAR
	func_block.IN1 := IN1;
	func_block.IN2 := IN2;
	func_block.IN3 := IN3;
	func_block.IN4 := IN4;
	func_block.IN5 := IN5;
	func_block.IN6 := IN6;
	func_block.IN7 := IN7;
	func_block.IN8 := IN8;
	func_block.X := X;

	func_block();
  	OUT1  := func_block.OUT1;
	OUT2  := func_block.OUT2;
	OUT3  := func_block.OUT3;
	OUT4  := func_block.OUT4;
	OUT5  := func_block.OUT5;
	OUT6  := func_block.OUT6;
	OUT7  := func_block.OUT7;
	OUT8  := func_block.OUT8;
	ID  := func_block.ID;
	X  := func_block.X;
END_PROGRAM

CONFIGURATION Config0
	RESOURCE Res0 ON PLC
		TASK task0(INTERVAL := T#20ms,PRIORITY := 0);
		PROGRAM instance0 WITH task0 : program0;
	END_RESOURCE
END_CONFIGURATION

(* ---- 661-ACTUATOR_A.ST ---- *)
FUNCTION_BLOCK T_PLC_MS_block
	VAR_OUTPUT
		T_PLC_MS :	UDINT;
	END_VAR

	VAR_EXTERNAL
		PLC_TICKS_PER_SEC :	INT;
		PLC_SYS_TICK_CNT :	DINT;
	END_VAR

	VAR
		debug :	BOOL;(*Debug-Mode ON / OFF*)
		N :	INT;(*Debug-Faktor*)
		Offset :	UDINT;(*Debug-Offset*)
		temp :	DWORD := DWORD#1;(*Debug-Offset*)
		mode :	BOOL;(*modus*)
		faktor :	UDINT;(*Systemtakt-Faktor*)
		init :	BOOL;
		v_plc_ticks_per_sec :	UDINT;
		base :	UDINT := UDINT#1000;
	END_VAR

	IF init = FALSE THEN
		v_plc_ticks_per_sec := INT_TO_UDINT(PLC_TICKS_PER_SEC);
		IF v_plc_ticks_per_sec = UDINT#1024 THEN
			faktor := UDINT#1;
			mode := FALSE;
		ELSIF v_plc_ticks_per_sec > UDINT#0 THEN
			IF v_plc_ticks_per_sec <= base THEN
				faktor := base / v_plc_ticks_per_sec;
				mode := FALSE;
			ELSE
				faktor := v_plc_ticks_per_sec / base;
				mode := TRUE;
			END_IF;
		ELSE
			faktor := UDINT#1;
		END_IF;
		init := TRUE;
	END_IF;

	IF mode THEN
		T_PLC_MS := DINT_TO_UDINT(PLC_SYS_TICK_CNT) / faktor;
	ELSE
		T_PLC_MS := DINT_TO_UDINT(PLC_SYS_TICK_CNT) * faktor;
	END_IF;

	IF debug THEN
		T_PLC_MS := (DWORD_TO_UDINT(SHL(UDINT_TO_DWORD(T_PLC_MS),N) OR SHL(temp,N)) - UDINT#1) + Offset;
	END_IF;

END_FUNCTION_BLOCK

FUNCTION_BLOCK CYCLE_4

	VAR_INPUT
		E :	BOOL := TRUE;
		T0 :	TIME;
		T1 :	TIME;
		T2 :	TIME;
		T3 :	TIME;
		S0 :	BOOL;
		SX :	INT;
		SL :	BOOL;
	END_VAR

	VAR_OUTPUT
		STATE :	INT;
	END_VAR

	VAR
		tx :	TIME;
		last :	TIME;
		init :	BOOL;
		T_PLC_MS :	T_PLC_MS_block;
	END_VAR

	T_PLC_MS();
	tx:= UDINT_TO_TIME(T_PLC_MS.T_PLC_MS);

	(* init on first cycle *)
	IF NOT init THEN
		init := TRUE;
		last := tx;
	END_IF;

	IF E THEN
		IF SL THEN
			(* when sx > 0 then the state sx is forced to start *)
			state:= LIMIT(0,SX,3);
			last := tx;
			(* this is to avoid to reset sx from the calling programm it does work fine on codesys but i am not sure about other systems, because we are writing to an input *)
			SL := FALSE;
		ELSE
			CASE state OF
				0 :	(* wait for T0 and switch to next cycle *)
					IF tx - last >= T0 THEN
						state := 1;
						last := tx;
					END_IF;
				1 : (* wait for T1 over 1st cycle *)
					IF tx - last >= T1 THEN
						state := 2;
						last := tx;
					END_IF;
				2 : (* wait for T1 over 1st cycle *)
					IF tx - last >= T2 THEN
						state := 3;
						last := tx;
					END_IF;
				3 : (* wait for T2 over 2nd cycle *)
					IF tx - last >= T3 THEN
						IF S0 THEN State := 0; END_IF; (* if S0 is false, the sequence stops at state 3 *)
						last := tx;
					END_IF;
			END_CASE;
		END_IF;
	ELSE
		state := 0;
		last := tx;
	END_IF;

END_FUNCTION_BLOCK

FUNCTION_BLOCK ACTUATOR_A_Block

	VAR_INPUT
		I1 :	BYTE;
		IS :	BOOL;
		I2 :	BYTE;
		RV :	BOOL;
		DX :	BOOL;
		RUNTIME :	TIME;
		SELF_ACT_TIME :	TIME;
		OUT_MIN :	DWORD;
		OUT_MAX :	DWORD;
	END_VAR

	VAR_OUTPUT
		Y :	DWORD;
	END_VAR

	VAR
		timer :	CYCLE_4;
		dx_edge :	BOOL;
	END_VAR

	timer(T0 := RUNTIME, T1 := RUNTIME, T3 := SELF_ACT_TIME, sl := DX AND NOT dx_edge, sx := 0, S0 := SELF_ACT_TIME > t#0s);
	dx_edge := dx;

	CASE timer.STATE OF
		0:
			Y := OUT_MIN;
		1:
			Y := OUT_MAX;
		3:
			IF rv THEN
				Y := UDINT_TO_DWORD(DWORD_TO_UDINT(OUT_MAX) - (DWORD_TO_UDINT(OUT_MAX) - DWORD_TO_UDINT(OUT_MIN)) * BYTE_TO_UDINT(SEL(IS, I1, I2)) / UDINT#255);
			ELSE
				Y := UDINT_TO_DWORD((DWORD_TO_UDINT(OUT_MAX) - DWORD_TO_UDINT(OUT_MIN)) * BYTE_TO_UDINT(SEL(IS, I1, I2)) / UDINT#255 + DWORD_TO_UDINT(OUT_MIN));
			END_IF;
	END_CASE;

END_FUNCTION_BLOCK

PROGRAM program0
	VAR
		I1 :	BYTE;
		IS :	BOOL;
		I2 :	BYTE;
		RV :	BOOL;
		DX :	BOOL;
		RUNTIME :	TIME;
		SELF_ACT_TIME :	TIME;
		OUT_MIN :	DWORD;
		OUT_MAX :	DWORD;
		Y :	DWORD;
		func_block : ACTUATOR_A_Block;
	END_VAR
	func_block.I1 := I1;
	func_block.IS := IS;
	func_block.I2 := I2 ;
	func_block.RV := RV;
	func_block.DX := DX;
	func_block.RUNTIME := RUNTIME;
	func_block.SELF_ACT_TIME := SELF_ACT_TIME ;
	func_block.OUT_MIN := OUT_MIN;
	func_block.OUT_MAX := OUT_MAX;
	func_block();
	Y  := func_block.Y;
END_PROGRAM

CONFIGURATION Config0
	VAR_GLOBAL
		PLC_TICKS_PER_SEC :	INT;
		PLC_SYS_TICK_CNT :	DINT;
	END_VAR
  	RESOURCE Res0 ON PLC
    	TASK task0(INTERVAL := T#20ms,PRIORITY := 0);
    	PROGRAM instance0 WITH task0 : program0;
  	END_RESOURCE
END_CONFIGURATION
